(* IEC 61131-3 sources: volt/packages/volt-lsp-iec/test-corpus/awa-palletizer/Device/Plc Logic/Application/Library Manager/L_TS2P_TechModulesSynchronizingCamming, 208 files *)

(* ---- L_MB1P_CLUTCHDIRECTION.dut ---- *)
TYPE L_MB1P_CLUTCHDIRECTION :
(
	MCNEGATIVEDIRECTION := -1,
	MCCURRENTDIRECTION := 0,
	MCPOSITIVEDIRECTION := 1
);
END_TYPE

(* ---- L_MB1P_CLUTCHMODE.dut ---- *)
TYPE L_MB1P_CLUTCHMODE :
(
	ABSOLUTE := 0,
	RELATIVE := 1,
	RAMP_POS := 2,
	RAMP_TIME := 3,
	RAMP_SLAVE_DIST := 4,
	ABSOLUTE_IN_TARGET := 5,
	RAMP_VELACC := 6,
	DISTRELATIVE := 7
);
END_TYPE

(* ---- L_MB1P_STATES.dut ---- *)
TYPE L_MB1P_STATES :
(
	INIT := 1,
	READY := 2,
	HOMING := 3,
	JOGGING := 10,
	JOGPOS := 11,
	JOGNEG := 12,
	POSITION_TRIMMING := 20,
	TRIM_POS_PLUS := 21,
	TRIM_POS_MINUS := 22,
	SYNCPOS := 30,
	POS_IS_SYNCHRONISED := 31,
	POSITIONING_TO_START_POS := 32,
	SYNCSPEED := 40,
	SPEED_IS_SYNCHRONISED := 41,
	DECOUPLED_LOCAL_DRIVING := 50,
	CONTMOTION := 60,
	PREPARING_PATH := 61,
	CHECK_LIMITS := 62,
	SYNCLINEVEL := 70,
	CAMMING := 80,
	CAMMING_DONE := 81,
	CLUTCH_OPEN_INSTANT := 82,
	CLUTCH_CLOSE := 83,
	CLUTCH_OPEN := 84,
	CYCLICMOTION := 130,
	SETPARAMETERS := 140,
	CAMSEQUENCER_LOADCAMTABLE := 150,
	CAMSEQUENCER_CYCLICCAM1 := 151,
	CAMSEQUENCER_CYCLICCAM3 := 152,
	CAMSEQUENCER_CAM1CYCLICCAM3CAM1 := 153,
	CAMSEQUENCER_CAM1CAM2CYCLICCAM3CAM4CAM1 := 154,
	CALCULATION := 798,
	BUSY := 799,
	DONE := 800,
	EMERGENCYSTOP := 991,
	SLOWSTOP := 992,
	ABC := 993,
	STANDBY := 994,
	HALT := 995,
	STOP := 996,
	QUICKSTOP := 997,
	SERVICE := 998,
	ERROR := 999,
	SYSTEMFAULT := 1000
);
END_TYPE

(* ---- L_TF1P_STATES.dut ---- *)
TYPE L_TF1P_STATES :
(
	INIT := 1,
	READY := 2,
	HOMING := 3,
	JOGGING := 10,
	JOGPOS := 11,
	JOGNEG := 12,
	POSITION_TRIMMING := 20,
	TRIM_POS_PLUS := 21,
	TRIM_POS_MINUS := 22,
	SYNCPOS := 30,
	POS_IS_SYNCHRONISED := 31,
	POSITIONING_TO_START_POS := 32,
	SYNCSPEED := 40,
	SPEED_IS_SYNCHRONISED := 41,
	DECOUPLED_LOCAL_DRIVING := 50,
	CONTMOTION := 60,
	PREPARING_PATH := 61,
	CHECK_LIMITS := 62,
	SYNCLINEVEL := 70,
	CAMMING := 80,
	CAMMING_DONE := 81,
	CLUTCH_OPEN_INSTANT := 82,
	CLUTCH_CLOSE := 83,
	CLUTCH_OPEN := 84,
	CYCLICMOTION := 130,
	SETPARAMETERS := 140,
	CAMSEQUENCER_LOADCAMTABLE := 150,
	CAMSEQUENCER_CYCLICCAM1 := 151,
	CAMSEQUENCER_CYCLICCAM3 := 152,
	CAMSEQUENCER_CAM1CYCLICCAM3CAM1 := 153,
	CAMSEQUENCER_CAM1CAM2CYCLICCAM3CAM4CAM1 := 154,
	STANDBY := 994,
	HALT := 995,
	STOP := 996,
	QUICKSTOP := 997,
	SERVICE := 998,
	ERROR := 999
);
END_TYPE

(* ---- L_TF1P_SYNCMODE.dut ---- *)
TYPE L_TF1P_SYNCMODE :
(
	ABSOLUTE := 0,
	RELATIVE := 1,
	RAMP_TIME := 3,
	RAMP_VELACC := 4,
	RAMP_DIST := 5,
	DISTRELATIVE := 7
);
END_TYPE

(* ---- L_TS2M_SCDATA_FLYINGSAWSTATE.dut ---- *)
TYPE L_TS2M_SCDATA_FLYINGSAWSTATE :
STRUCT
	XEXECUTEMOVETOPARKPOS : BOOL;
	XMOVETOPARKPOSBUSY : BOOL;
	XMOVETOPARKPOSDONE : BOOL;
	XMOVETOPARKPOSABORTED : BOOL;
	EMOVETOPARKPOSDIRECTION : MC_DIRECTION := MC_DIRECTION.mcPositiveDirection;
	XPARKPOSREACHED : BOOL;
	XINPARKPOSITION : BOOL;
	XSTARTFLYINGSAW : BOOL;
	XFMFLYINGSAWPOSITIONING : BOOL;
	XFMFLYINGSAWINPOSITION : BOOL;
	XFMERROR : BOOL;
	EFMERRORID : L_IE1P_Error;
	EFM_STATE : L_TB2P_States;
	LRSETACCELERATION : LREAL;
	LRSETVELOCITY : LREAL;
	LRSETPOSITION : LREAL;
END_STRUCT
END_TYPE

(* ---- L_TS2M_SCDATA_FM_FLYINGSAW.dut ---- *)
TYPE L_TS2M_SCDATA_FM_FLYINGSAW :
STRUCT
	LRSTARTPOSOUT : LREAL;
	XGETNEXTMARK : BOOL;
	XRESETGETNEXTMARK : BOOL;
	XRESETMARKSTACK : BOOL;
	XNEWMARKRECEIVED : BOOL;
	XMARKSTACKEMPTY : BOOL;
	XMARKVALID : BOOL;
	LRMARKPOSOUT : LREAL;
	POSPROFILERCLUTCH_XENABLE : BOOL;
	POSPROFILERCLUTCH_XSYNCVEL : BOOL;
	POSPROFILERCLUTCH_XSYNCPOS : BOOL;
	POSPROFILERCLUTCH_XSYNCOUTINSTANT : BOOL;
	POSPROFILERCLUTCH_XMOVETOTARGETPOS : BOOL;
	POSPROFILERCLUTCH_LRTARGETPOS : LREAL;
	POSPROFILERCLUTCH_LRCORRECTTIMEBASE : LREAL;
	POSPROFILERCLUTCH_XEXECUTEGAP : BOOL;
	POSPROFILERCLUTCH_XAUXEXECUTEGAP : BOOL;
	POSPROFILERCLUTCH_LRCYCMASTERPOS : LREAL;
	POSPROFILERCLUTCH_LRCYCMASTERVEL : LREAL;
	POSPROFILERCLUTCH_LRCYCMASTERACC : LREAL;
	POSPROFILERCLUTCH_XERROR : BOOL;
	POSPROFILERCLUTCH_XBUSY : BOOL;
	POSPROFILERCLUTCH_XDONE : BOOL;
	POSPROFILERCLUTCH_XACCDECSYNC : BOOL;
	POSPROFILERCLUTCH_XVELSYNCHRONISED : BOOL;
	POSPROFILERCLUTCH_XPOSSYNCHRONISED : BOOL;
	POSPROFILERCLUTCH_XPOSITIONING : BOOL;
	POSPROFILERCLUTCH_XINPOSITION : BOOL;
	POSPROFILERCLUTCH_LRSETSLAVEPOSOUT : LREAL;
	POSPROFILERCLUTCH_LRSETSLAVEVELOUT : LREAL;
	POSPROFILERCLUTCH_LRSETSLAVEACCOUT : LREAL;
	POSPROFILERCLUTCH_XPROFILERESETTIMEVALID : BOOL;
	POSPROFILERCLUTCH_LRPROFILERESETTIME : LREAL;
	XMODECHANGE : BOOL;
	EFLYINGSAWMODE_OLD : L_TS2P_FlyingSawMode;
	LRACCDIST : LREAL;
	LRACCTIME : LREAL;
	XTPRECEIVED : BOOL;
	LRTPACTPOSITION : LREAL;
	XMASTERITFVALID : BOOL;
	BYMASTERID : POINTER TO BYTE;
	XMASTERITFVALID_LOCK : BOOL;
	BYMASTERID_LOCK : POINTER TO BYTE;
	XWARNING_TPRECPOSITIONNOTSUPPORTED : BOOL;
	LRSYNCOUTPOS : LREAL;
	XSTATESAWSYNCHRONIZED : BOOL;
	XSYNCOVERRIDEACTIVE : BOOL;
	XRAMPGENBUSY : BOOL;
	LRCUTLENGTHPROCESSED : LREAL;
	LRDISTTOCUTPOSITION : LREAL;
	LRMASTERPOS1 : LREAL;
	LRMASTERPOS2 : LREAL;
	LRSLAVEPOS1 : LREAL;
	LRSLAVEPOS2 : LREAL;
	LRCUTGAP_INT : LREAL;
	XHEADCUTDONE : BOOL;
	XMOVETOLOWERLIMITBUSY : BOOL;
	LRDIST_INT : LREAL;
	XTIMESYNCINVALID : BOOL;
	LRTIMESYNCIN_INT : LREAL;
	XWAITINGFORNEXTCUTBUSY : BOOL;
	XBALANCEDPROFILEACTIVE : BOOL;
	LRDISTTOTARGET : LREAL;
	LRFILTMATERIALVEL : LREAL;
	LRFILTMATERIALACC : LREAL;
	LRRESTTIMETARGETTOLOWERLIMIT : LREAL;
	FB_STACKCONTROLARRAYNOISE : L_MC1P_StackControlArray := STRUCT(iMaxLegth := 10);
	ALRDELTAVEL : ARRAY [0..10] OF LREAL;
	AXNOISE : ARRAY [0..5] OF BOOL;
	ALRVELTOLERANCE : ARRAY [0..5] OF LREAL;
	XNOISE : BOOL;
	XACCPOSITIV : BOOL;
	IACCCHANGEDIRECTIONCOUNTER : INT;
	LRVELTOLERANCE_INT : LREAL;
	LRMAXVELTOLERANCE : LREAL;
	LRMAXACCTOLERANCE : LREAL;
	LRCYCMASTERVEL : LREAL;
	LRCYCMASTERVEL_OLD : LREAL;
END_STRUCT
END_TYPE

(* ---- L_TS2P_CAMDATAXYVA.dut ---- *)
TYPE L_TS2P_CAMDATAXYVA :
STRUCT
	LRX : LREAL;
	LRY : LREAL;
	LRYS : LREAL;
	LRYSS : LREAL;
	LRYSSS : LREAL;
END_STRUCT
END_TYPE

(* ---- L_TS2P_CAMSEQUENCEMODE.dut ---- *)
TYPE L_TS2P_CAMSEQUENCEMODE :
(
	CYCLICCAM1 := 0,
	CYCLICCAM3 := 1,
	CAM1_CYCLICCAM3_CAM1 := 2,
	CAM1_CAM2_CYCLICCAM3_CAM4_CAM1 := 3
);
END_TYPE

(* ---- L_TS2P_CAMSTOPMODE.dut ---- *)
TYPE L_TS2P_CAMSTOPMODE :
(
	HALT := 0,
	MOVETOPARKPOS := 1
);
END_TYPE

(* ---- L_TS2P_CLUTCHINMODE.dut ---- *)
TYPE L_TS2P_CLUTCHINMODE :
(
	DISTABSOLUTE := 2,
	INSTANTABSOLUTE := 10
);
END_TYPE

(* ---- L_TS2P_CLUTCHOUTMODE.dut ---- *)
TYPE L_TS2P_CLUTCHOUTMODE :
(
	DISTABSOLUTE := 2,
	DISTRELATIVE := 3
);
END_TYPE

(* ---- L_TS2P_CORRECTIONMODE.dut ---- *)
TYPE L_TS2P_CORRECTIONMODE :
(
	POLYNOM5TH := 0,
	PROFILEGENERATOR := 1
);
END_TYPE

(* ---- L_TS2P_COUPLINGMODE.dut ---- *)
TYPE L_TS2P_COUPLINGMODE :
(
	UNITCOUPLING := 0,
	COUPLINGOVERCYCLELENGTH := 1
);
END_TYPE

(* ---- L_TS2P_CROSSCUTTERSTATEIN.dut ---- *)
TYPE L_TS2P_CROSSCUTTERSTATEIN :
STRUCT
	MASTERVALUES : L_MC1P_IAXIS_REF_MASTERVALUES;
	XEXECUTEMOVETOPARKPOS : BOOL;
	XSYNCIN : BOOL;
	XHOLDINPARKPOS : BOOL;
	LRPRODUCTLENGTH : LREAL;
	LROVERSPEED : LREAL;
	LRSETOFFSETPOSX : LREAL;
	XTRIMPOS : BOOL;
	XTRIMNEG : BOOL;
	XTRIMRESET : BOOL;
	SCTPRECDATA_MARKSENSOR : L_MC1P_TpReceiveData;
	SCTPRECDATA_TOOLSENSOR : L_MC1P_TpReceiveData;
	XTEACHMARKWINDOW : BOOL;
	XTEACHMARKWINDOWTOOL : BOOL;
	XGEARFACTORCORR : BOOL;
	XGEARFACTORCORRHOLD : BOOL;
END_STRUCT
END_TYPE

(* ---- L_TS2P_CROSSCUTTERSTATEOUT.dut ---- *)
TYPE L_TS2P_CROSSCUTTERSTATEOUT :
STRUCT
	XSYNCHRONISED : BOOL;
	XACCDECSYNC : BOOL;
	XOFFSETTRIMACTIVE : BOOL;
	XINPARKPOS : BOOL;
	XHOLDINPARKPOSACTIVE : BOOL;
	XCUTDONE : BOOL;
	XCUTTINGACTIVE : BOOL;
	LRACTCUTLENGTH : LREAL;
	LROFFSETTOTAL : LREAL;
	XTRQCTRLACTIVE : BOOL;
	LRSETMARKCORROUT : LREAL;
	XMARKWINDOWTEACHED : BOOL;
	LRGEARFACTORCORR : LREAL;
	LRSETTOOLCORROUT : LREAL;
	XMARKWINDOWTEACHEDTOOL : BOOL;
END_STRUCT
END_TYPE

(* ---- L_TS2P_CUTTINGMODEBASE.dut ---- *)
TYPE L_TS2P_CUTTINGMODEBASE :
(
	CUT_LENGTH := 0,
	FLOW_PACKER := 1
);
END_TYPE

(* ---- L_TS2P_CUTTINGMODESTATE.dut ---- *)
TYPE L_TS2P_CUTTINGMODESTATE :
(
	CUT_LENGTH := 0,
	FLOW_PACKER := 1,
	CUT_LENGTH_TP_CORRECTION := 2,
	CUT_ON_TP := 3
);
END_TYPE

(* ---- L_TS2P_ELECTRONICGEARBOXBASEIN.dut ---- *)
TYPE L_TS2P_ELECTRONICGEARBOXBASEIN :
STRUCT
	MASTERVALUES : L_MC1P_IAXIS_REF_MASTERVALUES;
	XSYNCIN : BOOL;
	LRSETBASEVEL : LREAL;
	LRSETOFFSETPOS : LREAL;
	LRSETOFFSETVEL : LREAL;
	XTRIMPOS : BOOL;
	XTRIMNEG : BOOL;
	XTRIMRESET : BOOL;
	XINVERTGEARFACTOR : BOOL;
END_STRUCT
END_TYPE

(* ---- L_TS2P_ELECTRONICGEARBOXBASEOUT.dut ---- *)
TYPE L_TS2P_ELECTRONICGEARBOXBASEOUT :
STRUCT
	XSYNCHRONISED : BOOL;
	XACCDECSYNC : BOOL;
	XOFFSETTRIMACTIVE : BOOL;
	XBASEVELOCITYACTIVE : BOOL;
	LROFFSETTOTALVEL : LREAL;
END_STRUCT
END_TYPE

(* ---- L_TS2P_FLEXCAMHIGHIN.dut ---- *)
TYPE L_TS2P_FLEXCAMHIGHIN :
STRUCT
	MASTERVALUES : L_MC1P_IAXIS_REF_MASTERVALUES;
	XCLUTCHCLOSE : BOOL;
	XLOADCLUTCHPOS : BOOL;
	LRLOADCLUTCHPOS : LREAL;
	XFINDCLUTCHXPOS : BOOL;
	XSYNCIN : BOOL;
	XSYNCPOSRESTORE : BOOL;
	XCAMCHANGEINSTANT : BOOL;
	LRSETOFFSETPOSX : LREAL;
	LRSETOFFSETPOSY : LREAL;
	LRSETSCALINGX : LREAL;
	LRSETSCALINGY : LREAL;
	CAMTABLE1 : MC_CAM_REF;
	CAMTABLE2 : MC_CAM_REF;
	CAMTABLE3 : MC_CAM_REF;
	CAMTABLE4 : MC_CAM_REF;
	WSETCAMTABLE : WORD := 1;
	XCAMSEQUENCER : BOOL;
END_STRUCT
END_TYPE

(* ---- L_TS2P_FLEXCAMHIGHOUT.dut ---- *)
TYPE L_TS2P_FLEXCAMHIGHOUT :
STRUCT
	XCLUTCHACTIVE : BOOL;
	XCLUTCHCLOSED : BOOL;
	XACCDECSYNC : BOOL;
	XSYNCHRONISED : BOOL;
	XMOVETOPARKPOSACTIVE : BOOL;
	XINPARKPOS : BOOL;
	XENDOFPROFILE : BOOL;
	LROFFSETPOSX : LREAL;
	LROFFSETPOSY : LREAL;
	LROFFSETSYNCPOS : LREAL;
	WACTIVECAMTABLE : WORD;
	XCAMSEQUENCERACTIVE : BOOL;
END_STRUCT
END_TYPE

(* ---- L_TS2P_FLEXCAMSTATEIN.dut ---- *)
TYPE L_TS2P_FLEXCAMSTATEIN :
STRUCT
	MASTERVALUES : L_MC1P_IAXIS_REF_MASTERVALUES;
	XSYNCIN : BOOL;
	XCAMCHANGEINSTANT : BOOL;
	LRSETOFFSETPOSX : LREAL;
	LRSETOFFSETPOSY : LREAL;
	LRSETSCALINGX : LREAL := 1;
	LRSETSCALINGY : LREAL := 1;
	CAMTABLE1 : MC_CAM_REF;
	CAMTABLE2 : MC_CAM_REF;
	CAMTABLE3 : MC_CAM_REF;
	CAMTABLE4 : MC_CAM_REF;
	WSETCAMTABLE : WORD := 1;
	XCAMSEQUENCER : BOOL;
END_STRUCT
END_TYPE

(* ---- L_TS2P_FLEXCAMSTATEOUT.dut ---- *)
TYPE L_TS2P_FLEXCAMSTATEOUT :
STRUCT
	XSYNCHRONISED : BOOL;
	XACCDECSYNC : BOOL;
	XCAMMINGBUSY : BOOL;
	XENDOFPROFILE : BOOL;
	LROFFSETPOSX : LREAL;
	LROFFSETPOSY : LREAL;
	WACTIVECAMTABLE : WORD;
	XCAMSEQUENCERACTIVE : BOOL;
END_STRUCT
END_TYPE

(* ---- L_TS2P_FLYINGSAWMODE.dut ---- *)
TYPE L_TS2P_FLYINGSAWMODE :
(
	MARKCONTROLLED := 0,
	LENGTHCONTROLLED := 1,
	LENGTHCONTROLLEDAUTOSYNC := 2
);
END_TYPE

(* ---- L_TS2P_FLYINGSAWPROFILEMODE.dut ---- *)
TYPE L_TS2P_FLYINGSAWPROFILEMODE :
(
	DEFAULT := 0,
	BALANCED := 1
);
END_TYPE

(* ---- L_TS2P_FLYINGSAWSTATEIN.dut ---- *)
TYPE L_TS2P_FLYINGSAWSTATEIN :
STRUCT
	MASTERVALUES : L_MC1P_IAXIS_REF_MASTERVALUES;
	XSTARTFLYINGSAW : BOOL;
	XSYNCININSTANT : BOOL;
	XEXECUTENEXTCUT : BOOL;
	XEXECUTEGAP : BOOL;
	XSETCUTTINGLENGTHINSTANT : BOOL;
	LRCUTTINGLENGTH : LREAL;
	LRSYNCOVERRIDE : LREAL := 1;
	XSETMATERIALCOUNTER : BOOL;
	XMOVETOPARKPOS : BOOL;
	XRESUMETARGETPOS : BOOL;
	XRESETMARKSTACK : BOOL;
	SCTPRECDATA_MARKSENSOR : L_MC1P.L_MC1P_TpReceiveData;
END_STRUCT
END_TYPE

(* ---- L_TS2P_FLYINGSAWSTATEOUT.dut ---- *)
TYPE L_TS2P_FLYINGSAWSTATEOUT :
STRUCT
	XSYNCHRONISED : BOOL;
	XACCDECSYNC : BOOL;
	XINPOSITION : BOOL;
	XPOSITIONING : BOOL;
	LRMATERIALCOUNTER : LREAL;
	LRTARGETPOS : LREAL;
	LRCUTGAP : LREAL;
	LRACTIVECUTTINGLENGTH : LREAL;
	WMARKSINSTACK : WORD;
END_STRUCT
END_TYPE

(* ---- L_TS2P_FLYINGSAWSTOPMODE.dut ---- *)
TYPE L_TS2P_FLYINGSAWSTOPMODE :
(
	HALT := 0,
	MOVETOPARKPOS := 1
);
END_TYPE

(* ---- L_TS2P_INTERFACEID.dut ---- *)
TYPE L_TS2P_INTERFACEID :
(
	L_TS2P_ISTRUCTPROVIDERFLYINGSAW := (L_TS2P_Internal.cdiEnumStartValue + 1),
	L_TS2P_ISTRUCTPROVIDERSYNCPOS := (L_TS2P_Internal.cdiEnumStartValue + 2),
	L_TS2P_ISTRUCTPROVIDERSYNCANDCORRECTION := (L_TS2P_Internal.cdiEnumStartValue + 3),
	L_TS2P_ISTRUCTPROVIDERFLEXCAMHIGH := (L_TS2P_Internal.cdiEnumStartValue + 4)
);
END_TYPE

(* ---- L_TS2P_OFFSETMODE.dut ---- *)
TYPE L_TS2P_OFFSETMODE :
(
	X_ZERO := 0,
	INSTANTABSOLUTE := 1,
	PROFGENABSOLUTE := 2
);
END_TYPE

(* ---- L_TS2P_SCALINGMODE.dut ---- *)
TYPE L_TS2P_SCALINGMODE :
(
	X_ZERO := 0,
	INSTANTABSOLUTE := 1,
	INSTANTRELATIVE := 2,
	PROFGENABSOLUTE := 3,
	PROFGENRELATIVE := 4
);
END_TYPE

(* ---- L_TS2P_SCAP_CROSSCUTTERBASE.dut ---- *)
TYPE L_TS2P_SCAP_CROSSCUTTERBASE :
STRUCT
END_STRUCT
END_TYPE

(* ---- L_TS2P_SCAP_CROSSCUTTERHIGH.dut ---- *)
TYPE L_TS2P_SCAP_CROSSCUTTERHIGH :
STRUCT
END_STRUCT
END_TYPE

(* ---- L_TS2P_SCAP_CROSSCUTTERSTATE.dut ---- *)
TYPE L_TS2P_SCAP_CROSSCUTTERSTATE :
STRUCT
END_STRUCT
END_TYPE

(* ---- L_TS2P_SCAP_ELECTRONICGEARBOXBASE.dut ---- *)
TYPE L_TS2P_SCAP_ELECTRONICGEARBOXBASE :
STRUCT
END_STRUCT
END_TYPE

(* ---- L_TS2P_SCAP_FLEXCAMHIGH.dut ---- *)
TYPE L_TS2P_SCAP_FLEXCAMHIGH :
STRUCT
END_STRUCT
END_TYPE

(* ---- L_TS2P_SCAP_FLEXCAMSTATE.dut ---- *)
TYPE L_TS2P_SCAP_FLEXCAMSTATE :
STRUCT
END_STRUCT
END_TYPE

(* ---- L_TS2P_SCAP_FLYINGSAWSTATE.dut ---- *)
TYPE L_TS2P_SCAP_FLYINGSAWSTATE :
STRUCT
END_STRUCT
END_TYPE

(* ---- L_TS2P_SCAP_SYNCANDCORRECTIONSTATE.dut ---- *)
TYPE L_TS2P_SCAP_SYNCANDCORRECTIONSTATE :
STRUCT
END_STRUCT
END_TYPE

(* ---- L_TS2P_SCAP_SYNCPOSBASE.dut ---- *)
TYPE L_TS2P_SCAP_SYNCPOSBASE :
STRUCT
END_STRUCT
END_TYPE

(* ---- L_TS2P_SCAP_TM_CROSSCUTTERBASE.dut ---- *)
TYPE L_TS2P_SCAP_TM_CROSSCUTTERBASE :
STRUCT
	AP_XENDOFPROFILEWINDOWSIZE : BOOL;
	AP_LRENDOFPROFILEWINDOWSIZE : LREAL := 0;
	AP_XOVERSPEEDUPPERLIMIT : BOOL;
	AP_LROVERSPEEDUPPERLIMIT : LREAL := 2;
	AP_XSETOFFSETSLAVE : BOOL;
	AP_LRSETOFFSETSLAVE : LREAL;
	AP_XOFFSETSLAVEPAR : BOOL;
	AP_LROFFSETSLAVEVEL : LREAL;
	AP_LROFFSETSLAVEACC : LREAL;
	AP_LROFFSETSLAVEDEC : LREAL;
	AP_LROFFSETSLAVEJERK : LREAL;
END_STRUCT
END_TYPE

(* ---- L_TS2P_SCAP_TM_CROSSCUTTERHIGH.dut ---- *)
TYPE L_TS2P_SCAP_TM_CROSSCUTTERHIGH :
STRUCT
END_STRUCT
END_TYPE

(* ---- L_TS2P_SCAP_TM_CROSSCUTTERSTATE.dut ---- *)
TYPE L_TS2P_SCAP_TM_CROSSCUTTERSTATE :
STRUCT
	AP_XTPAXISDELAYCYCLE : BOOL;
	AP_LRTPAXISDELAYCYCLE : LREAL;
	AP_XTPAXISCOMPFACTOR : BOOL;
	AP_LRTPAXISCOMPFACTOR : LREAL;
	AP_XUPPERCORRPOS : BOOL;
	AP_LRUPPERCORRPOS : LREAL;
	AP_XLOWERCORRPOS : BOOL;
	AP_LRLOWERCORRPOS : LREAL;
	AP_XCUTTINGANGLESTOPCAM : BOOL;
	AP_LRCUTTINGANGLESTOPCAM : LREAL := 10;
	AP_XSETCUTLENGTHINPRODUCT : BOOL;
END_STRUCT
END_TYPE

(* ---- L_TS2P_SCAP_TM_ELECTRONICGEARBOXBASE.dut ---- *)
TYPE L_TS2P_SCAP_TM_ELECTRONICGEARBOXBASE :
STRUCT
	AP_XGEARINGNUMERATOR : BOOL;
	AP_DWGEARINGNUMERATOR : DWORD := 1;
	AP_XGEARINGDENOMINATOR : BOOL;
	AP_DWGEARINGDENOMINATOR : DWORD := 1;
	AP_XLIMITALLOWEDDIRECTION : BOOL;
	AP_LREXTTHRESHOLDDIRECTION : LREAL;
END_STRUCT
END_TYPE

(* ---- L_TS2P_SCAP_TM_FLEXCAM.dut ---- *)
TYPE L_TS2P_SCAP_TM_FLEXCAM :
STRUCT
	AP_LREXTTHRESHOLDDIRECTION : LREAL;
	AP_LRMASTERVELSTANDSTILLDEADBAND : LREAL;
	AP_XENDOFPROFILEWINDOWSIZE : BOOL;
	AP_LRENDOFPROFILEWINDOWSIZE : LREAL;
	AP_XSETVALUEMODE : BOOL;
	AP_ESETVALUEMODE : L_MC1P_SetValueMode := L_MC1P_SetValueMode.PosVelAcc;
END_STRUCT
END_TYPE

(* ---- L_TS2P_SCAP_TM_FLEXCAMBASE.dut ---- *)
TYPE L_TS2P_SCAP_TM_FLEXCAMBASE :
STRUCT
	AP_XENDOFPROFILEWINDOWSIZE : BOOL;
	AP_LRENDOFPROFILEWINDOWSIZE : LREAL := 0;
	AP_XCALCAMPROFILER : BOOL := TRUE;
	AP_XSETVALUEMODE : BOOL;
	AP_ESETVALUEMODE : L_MC1P_SetValueMode := L_MC1P_SetValueMode.PosVelAcc;
END_STRUCT
END_TYPE

(* ---- L_TS2P_SCAP_TM_FLEXCAMSTATE.dut ---- *)
TYPE L_TS2P_SCAP_TM_FLEXCAMSTATE :
STRUCT
END_STRUCT
END_TYPE

(* ---- L_TS2P_SCAP_TM_FLYINGSAWSTATE.dut ---- *)
TYPE L_TS2P_SCAP_TM_FLYINGSAWSTATE :
STRUCT
	AP_XLOADTOTALCUTTINGLENGTH : BOOL;
	AP_LRLOADTOTALCUTTINGLENGTH : LREAL;
	AP_XLOADTARGETPOS : BOOL;
	AP_LRLOADTARGETPOS : LREAL;
	AP_XRANGEOFTOLERANCE : BOOL;
	AP_LRRANGEOFTOLERANCE : LREAL;
	AP_XMARKDETECTERRCOMP : BOOL;
	AP_LRMARKDETECTERRCOMP : LREAL;
	AP_XTASKCYCLEDELAY : BOOL;
	AP_BYTASKCYCLEDELAY : BYTE;
END_STRUCT
END_TYPE

(* ---- L_TS2P_SCAP_TM_SYNCANDCORRECTIONSTATE.dut ---- *)
TYPE L_TS2P_SCAP_TM_SYNCANDCORRECTIONSTATE :
STRUCT
	AP_DIDEADTIMECOMP : DINT;
END_STRUCT
END_TYPE

(* ---- L_TS2P_SCAP_TM_SYNCPOSBASE.dut ---- *)
TYPE L_TS2P_SCAP_TM_SYNCPOSBASE :
STRUCT
	AP_XLOADGEARBOXPOSOUT : BOOL;
	AP_LRLOADGEARBOXPOSOUT : LREAL;
	AP_XLOADTRIMOFFSET : BOOL;
	AP_LRLOADTRIMOFFSET : LREAL;
	AP_XLOADOFFSETSYNC : BOOL;
	AP_LRLOADOFFSETSYNC : LREAL;
	AP_XLIMITALLOWEDDIRECTION : BOOL;
	AP_LREXTTHRESHOLDDIRECTION : LREAL;
	AP_LRMASTERVELSTANDSTILLDEADBAND : LREAL;
END_STRUCT
END_TYPE

(* ---- L_TS2P_SCDATA_TM_FLEXCAM.dut ---- *)
TYPE L_TS2P_SCDATA_TM_FLEXCAM :
STRUCT
	XEXECUTEMOVETOPARKPOS : BOOL;
	XHALTFLEXCAM : BOOL;
	XMOVETOPARKPOSBUSY : BOOL;
	XMOVETOPARKPOSABORTED : BOOL;
	MASTERVALUES_ITFVALID : L_MC1P_IAXIS_REF_MASTERVALUES;
	LRMASTERPOS_OLD : LREAL;
	LRMASTERVEL_OLD : LREAL;
	LRSETPOSITIONFORSYNCMASTER : LREAL;
	LRSETVELOCITYFORSYNCMASTER : LREAL;
	LRSETACCELERATIONFORSYNCMASTER : LREAL;
	LRCYCLELENGTHMASTER : LREAL;
	ETRAVERSINGRANGEMASTER : L_MC1P_TraversingRange;
	LRSETPOSITIONAXIS : LREAL;
	LRSETVELOCITYAXIS : LREAL;
	LRSETACCELERATIONAXIS : LREAL;
	WACTDIRECTIONMASTER : WORD;
	XCAMSEQUENCERERROR : BOOL;
	ECAMSEQUENCERERROR : L_IE1P_Error;
	XCAMERROR : BOOL;
	ECAMERROR : L_IE1P_Error;
	XCAMBUSY : BOOL;
	XCAMDONE : BOOL;
	XLOCKTOCAMRESTORE : BOOL;
	ESYNCINMODE : L_TS2P_SyncInMode := L_TS2P_SyncInMode.ProfGenAbsolute;
	XCLUTCHBUSY : BOOL;
	XCLUTCHDONE : BOOL;
	XCLUTCHACCDECSYNCLED : BOOL;
	LRSETCLUTCHPOSOUT : LREAL;
	LRSETCLUTCHVELOUT : LREAL;
	LRSETCLUTCHACCOUT : LREAL;
	LRSETCLUTCHPOSOUTOLD : LREAL;
	LRSETCLUTCHVELOUTOLD : LREAL;
	XCLUTCHERROR : BOOL;
	ECLUTCHERROR : L_IE1P_Error;
	XENABLEALLOWEDDIRECTION : BOOL;
	LRALLOWEDDIRECTIONSETPOSOUT : LREAL;
	LRALLOWEDDIRECTIONSETVELOUT : LREAL;
	LRALLOWEDDIRECTIONSETACCOUT : LREAL;
	XALLOWEDDIRECTIONERROR : BOOL;
	XALLOWEDDIRECTIONWARNING : BOOL;
	EALLOWEDDIRECTIONERROR : L_IE1P_Error;
	XPOSFOLLOWERENABLE : BOOL;
	XPOSFOLLOWERBUSY : BOOL;
	XENABLETRANSSYNCHRONISED : BOOL;
	LRTASKCYCLE : LREAL;
	XLOCKTOCAM : BOOL;
	XCAMCHANGEINSTANT_INT : BOOL;
	LRSETOFFSETMASTER_INT : LREAL;
	LRSETOFFSETSLAVE_INT : LREAL;
	LRSETSCALINGMASTER_INT : LREAL := 1;
	LRSETSCALINGSLAVE_INT : LREAL := 1;
	SCPAR_INT : L_TS2P_scPar_TM_FlexCam;
	XLOCKTOCAMERROR : BOOL;
	ELOCKTOCAMERROR : L_IE1P_Error;
	XCAMTABLEVALID : BOOL;
	XCAMMINGBUSY : BOOL;
	XLOCKTOCAMDONE : BOOL;
	XLOCKTOCAMBUSY : BOOL;
	XLOCKTOCAMBUSYLED : BOOL;
	XLOCKTOCAMBUSYGENERAL : BOOL;
	EPOSFOLLOWERMODE : L_MC1P_SetValueMode;
	XLOADCAMXVALUEBUSY : BOOL;
	XDIRECTIONLIMITED : BOOL;
	XFINDCLUTCHXPOS : BOOL;
	XVISULAMPFALSE : BOOL;
	LRSETVELOLD : LREAL;
END_STRUCT
END_TYPE

(* ---- L_TS2P_SCDATA_TM_SYNCANDCORRECTIONSTATE.dut ---- *)
TYPE L_TS2P_SCDATA_TM_SYNCANDCORRECTIONSTATE :
STRUCT
	MASTERVALUES_ITFVALID : L_MC1P_IAXIS_REF_MASTERVALUES;
	XMASTERITFVALID : BOOL;
	XMASTERVALUECORRENABLED : BOOL;
	LRSETPOSOLD : LREAL;
	LRMASTERSETPOSOLD : LREAL;
	LRMASTERACTPOSITIONOLD : LREAL;
	LRSETVELOCITYGEARING : LREAL;
	LRSENSORSETPOS : LREAL;
	XMARKDISTCHANGED : BOOL;
	LRACTOFFSETMASTER : LREAL;
	LRACTOFFSETSLAVE : LREAL;
	LRLOWERCORRPOS : LREAL;
	LRUPPERCORRPOS : LREAL;
	LRMARKDIST : LREAL;
	LRACTOFFSETX : LREAL;
	XVALUESTORED : BOOL;
	XFIRSTVALUESTORED : BOOL;
	XTEACHTPSENSOROLD : BOOL;
	XTPSENSORTEACHEDOLD : BOOL;
	LRMARKSTACKLENGTH : LREAL;
	DWACTTIMESTAMPMARKWINDOW : DWORD;
	DWRECTIMESTAMPMARKWINDOW : DWORD;
	XVALUESTOREDMARKWINDOW : BOOL;
	XSUPPORTTIMESTAMPMARKWINDOW : BOOL;
	XVALUESTOREDMARKSTACK : BOOL;
	DWACTTIMESTAMPMARKSTACK : DWORD;
	DWRECTIMESTAMPMARKSTACK : DWORD;
	XVALUESTOREDTPCONVERTER : BOOL;
	LRTPACTPOSITIONTPCONVERTER : LREAL;
	LRACTMARKDIST : LREAL;
	LRMARKDISTINTEGRATOR : LREAL;
	LRTPDEADTIMEDIFF : LREAL;
	LRMARKERROR : LREAL;
	LRMARKERRORLIMITED : LREAL;
	LRMARKERRORGEARFACTOR : LREAL;
	LRCORRRESIDUAL : LREAL;
	LRDELTAGEARFACTORCORR : LREAL;
	LRGEARFACTORINTEGRATOR : LREAL;
	LRGEARFACTORNUMERATOR : LREAL;
	LRGEARFACTORNUMERATORCORR : LREAL;
	LRGEARFACTORDENOMINATOR : LREAL;
	LRGEARFACTORNUMERATORCORRLIMITED : LREAL;
	LRSTARTPOS : LREAL;
	ECORRMODEMASTEROLD : L_TS2P_CorrectionMode;
	LRSETVELOUTCORRECTION : LREAL;
	LRSETPOSOUTCORRECTION : LREAL;
	XVALUESTOREDCORRMARKERROR : BOOL;
END_STRUCT
END_TYPE

(* ---- L_TS2P_SCDATA_TM_SYNCPOSBASE.dut ---- *)
TYPE L_TS2P_SCDATA_TM_SYNCPOSBASE :
STRUCT
	MASTERVALUES_ITFVALID : L_MC1P_IAXIS_REF_MASTERVALUES;
	XHOMINGNOTNEEDED : BOOL;
	LRSETPOSITIONFORSYNCMASTER : LREAL;
	LRSETVELOCITYFORSYNCMASTER : LREAL;
	LRSETACCELERATIONFORSYNCMASTER : LREAL;
	LRCYCLELENGTHMASTER : LREAL;
	ETRAVERSINGRANGEMASTER : L_MC1P_TraversingRange;
	WACTDIRECTIONMASTER : WORD;
	XOFFSETTRIMERROR : BOOL;
	EOFFSETTRIMERROR : L_IE1P_Error;
	XADDOFFSETERROR : BOOL;
	EADDOFFSETERROR : L_IE1P_Error;
	LROFFSETAXISCONVERTER : LREAL;
	WTRAVERSINGRANGECOMBINATION : WORD;
	WTRAVERSINGRANGECOMBINATIONOLD : WORD;
	XGEARBOXERROR : BOOL;
	EGEARBOXERROR : L_IE1P_Error;
	LRBASEVELLIMITED : LREAL;
	XCLUTCHENABLE : BOOL;
	XCLUTCHSYNCIN : BOOL;
	XCLUTCHSYNCPOSRESTORE : BOOL;
	LRSETVELCLUTCHOFFSET : LREAL;
	LRSETACCCLUTCHOFFSET : LREAL;
	LRSETDECCLUTCHOFFSET : LREAL;
	LRSETJERKCLUTCHOFFSET : LREAL;
	ESYNCMODE : L_TB2P_SyncMode := L_TB2P_SyncMode.ProfGenAbsolute;
	XCLUTCHBUSY : BOOL;
	XCLUTCHDONE : BOOL;
	XCLUTCHSYNCHRONISED : BOOL;
	XCLUTCHACCDECSYNC : BOOL;
	LRCLUTCHSETPOSOUT : LREAL;
	LRCLUTCHSETVELOUT : LREAL;
	LRCLUTCHSETACCOUT : LREAL;
	LRSYNCOFFSET : LREAL;
	XCLUTCHERROR : BOOL;
	ECLUTCHERROR : L_IE1P_Error;
	LRALLOWEDDIRECTIONSETPOSOUT : LREAL;
	LRALLOWEDDIRECTIONSETVELOUT : LREAL;
	LRALLOWEDDIRECTIONSETACCOUT : LREAL;
	XALLOWEDDIRECTIONERROR : BOOL;
	XALLOWEDDIRECTIONWARNING : BOOL;
	EALLOWEDDIRECTIONERROR : L_IE1P_Error;
	XPOSFOLLOWERENABLE : BOOL;
	LRPOSFOLLOWERSETPOSIN : LREAL;
	LRPOSFOLLOWERSETVELIN : LREAL;
	XENABLETRANSBASEVEL : BOOL;
	XENABLETRANSSYNCHRONISED : BOOL;
	XENABLEOLD : BOOL;
	LRTASKCYCLE : LREAL;
	LRCYCLELENGTH : LREAL;
	ETRAVERSINGRANGE : L_MC1P_TraversingRange;
	LRSETPOSITION : LREAL;
	LRSETVELOCITY : LREAL;
	LRSETACCELERATION : LREAL;
	XREQUESTTOSTANDBY : BOOL;
END_STRUCT
END_TYPE

(* ---- L_TS2P_SCERRORINFO.dut ---- *)
TYPE L_TS2P_SCERRORINFO :
STRUCT
	XERROR : BOOL;
	XWARNING : BOOL;
	EERRORID : L_IE1P_Error;
	XAXISERROR : BOOL;
	XAXISWARNING : BOOL;
	EAXISERRORID : L_IE1P_Error;
	XDRIVEERROR : BOOL;
	XDRIVEWARNING : BOOL;
	DWDRIVEERRORID : DWORD;
END_STRUCT
END_TYPE

(* ---- L_TS2P_SCPAR_CROSSCUTTERBASE.dut ---- *)
TYPE L_TS2P_SCPAR_CROSSCUTTERBASE :
STRUCT
END_STRUCT
END_TYPE

(* ---- L_TS2P_SCPAR_CROSSCUTTERSTATE.dut ---- *)
TYPE L_TS2P_SCPAR_CROSSCUTTERSTATE :
STRUCT
END_STRUCT
END_TYPE

(* ---- L_TS2P_SCPAR_ELECTRONICGEARBOXBASE.dut ---- *)
TYPE L_TS2P_SCPAR_ELECTRONICGEARBOXBASE :
STRUCT
END_STRUCT
END_TYPE

(* ---- L_TS2P_SCPAR_FLEXCAMHIGH.dut ---- *)
TYPE L_TS2P_SCPAR_FLEXCAMHIGH :
STRUCT
END_STRUCT
END_TYPE

(* ---- L_TS2P_SCPAR_FLEXCAMSTATE.dut ---- *)
TYPE L_TS2P_SCPAR_FLEXCAMSTATE :
STRUCT
END_STRUCT
END_TYPE

(* ---- L_TS2P_SCPAR_FLYINGSAWSTATE.dut ---- *)
TYPE L_TS2P_SCPAR_FLYINGSAWSTATE :
STRUCT
END_STRUCT
END_TYPE

(* ---- L_TS2P_SCPAR_SYNCANDCORRECTIONSTATE.dut ---- *)
TYPE L_TS2P_SCPAR_SYNCANDCORRECTIONSTATE :
STRUCT
END_STRUCT
END_TYPE

(* ---- L_TS2P_SCPAR_SYNCPOSBASE.dut ---- *)
TYPE L_TS2P_SCPAR_SYNCPOSBASE :
STRUCT
END_STRUCT
END_TYPE

(* ---- L_TS2P_SCPAR_TM_CROSSCUTTERBASE.dut ---- *)
TYPE L_TS2P_SCPAR_TM_CROSSCUTTERBASE :
STRUCT
	LRSETOFFSETTRIMVEL : LREAL := 10.0;
	LRSETOFFSETTRIMACC : LREAL := 100.0;
	LRSETOFFSETTRIMDEC : LREAL := 100.0;
	LRSETOFFSETTRIMJERK : LREAL := 10000.0;
	ETRIMMODE : L_TS2P_TrimMode := L_TS2P_TrimMode.position;
	LRTRIMDIST : LREAL := 1;
	ESYNCMODE : L_TS2P_SyncModeCrossCutter;
	LRMASTERSYNCINDIST : LREAL := 0;
	LRMASTERSYNCOUTDIST : LREAL := 0;
	XMASTERABSOLUTE : BOOL := TRUE;
	LRSTARTXPOSRELATIVE : LREAL := 0;
	BYSTARTTOOLNO : BYTE := 0;
	BYNUMOFTOOLS : BYTE := 1;
	LRCUTTINGANGLE : LREAL := 10;
	LRTOOLCIRCUMFERENCE : LREAL := 75.55555;
	XCALCCAMBOUNDS : BOOL := FALSE;
	LRMASTERMAXVEL : LREAL := 100;
	LRMASTERMAXACC : LREAL := 1000;
	LRSCALINGMASTER : LREAL := 1;
	EPROFILETYPE : L_MC2P_LawOfMotion := L_MC2P_LawOfMotion.Poly5;
END_STRUCT
END_TYPE

(* ---- L_TS2P_SCPAR_TM_CROSSCUTTERBASEEXTENSION.dut ---- *)
TYPE L_TS2P_SCPAR_TM_CROSSCUTTERBASEEXTENSION :
STRUCT
	ECUTTINGMODE : L_TS2P_CuttingModeBase := L_TS2P_CuttingModeBase.cut_length;
END_STRUCT
END_TYPE

(* ---- L_TS2P_SCPAR_TM_CROSSCUTTERHIGH.dut ---- *)
TYPE L_TS2P_SCPAR_TM_CROSSCUTTERHIGH :
STRUCT
END_STRUCT
END_TYPE

(* ---- L_TS2P_SCPAR_TM_CROSSCUTTERSTATE.dut ---- *)
TYPE L_TS2P_SCPAR_TM_CROSSCUTTERSTATE :
STRUCT
	ECUTTINGMODE : L_TS2P_CuttingModeState;
	ALRCUTLENGTHINPRODUCT : ARRAY [1..10] OF LREAL;
	LRMINPRODUCTLENGTH : LREAL := 50;
	LRTRQCTRLGAIN : LREAL := 0;
	LRTRQCTRLRATETIME : LREAL := 0;
	LRMINERTIA : LREAL := 0;
	XCORRMARKERRORMASTER : BOOL := TRUE;
	LRSENSORTOOLDISTMASTER : LREAL := 0.0;
	LRMAXCORRPOSMASTER : LREAL := 30.0;
	LRMAXCORRNEGMASTER : LREAL := -30.0;
	XENABLEMARKWINDOWMASTER : BOOL;
	LRMARKWINDOWSIZEMASTER : LREAL := 90.0;
	LRSETOFFSETMARKWINDOWMASTER : LREAL := 0.0;
	LRGEARFACTORCORRGAINMASTER : LREAL := 0.1;
	LRMAXGEARFACTORCORRMASTER : LREAL := 10;
	DWMAXNUMBERVIRTUALMARKSMASTER : DWORD := 5;
	XLOADREGPOS : BOOL;
	LRLOADREGPOS : LREAL;
	XCALCTOOLERROR : BOOL := FALSE;
	XCORRTOOLERROR : BOOL := TRUE;
	LRSENSORTOOLDISTTOOL : LREAL := 0.0;
	XENABLEMARKWINDOWTOOL : BOOL := FALSE;
	LRMAXCORRPOSTOOL : LREAL := 30.0;
	LRMAXCORRNEGTOOL : LREAL := -30.0;
	LRUPPERCORRPOSTOOL : LREAL := 180.0;
	LRLOWERCORRPOSTOOL : LREAL := 90.0;
	LRMARKWINDOWSIZETOOL : LREAL := 90.0;
	LRSETOFFSETMARKWINDOWTOOL : LREAL := 0.0;
	DWMAXNUMBERVIRTUALMARKSTOOL : DWORD := 5;
END_STRUCT
END_TYPE

(* ---- L_TS2P_SCPAR_TM_ELECTRONICGEARBOXBASE.dut ---- *)
TYPE L_TS2P_SCPAR_TM_ELECTRONICGEARBOXBASE :
STRUCT
	ECOUPLINGMODE : L_TS2P_CouplingMode := 1;
	LRTOLERANCEINVERTGEARFACTOR : LREAL := 0;
END_STRUCT
END_TYPE

(* ---- L_TS2P_SCPAR_TM_FLEXCAM.dut ---- *)
TYPE L_TS2P_SCPAR_TM_FLEXCAM :
STRUCT
	ECLUTCHINMODE : L_TS2P_ClutchInMode := L_TS2P_ClutchInMode.DistAbsolute;
	ECLUTCHOUTMODE : L_TS2P_ClutchOutMode := L_TS2P_ClutchOutMode.DistAbsolute;
	LRCLUTCHINDISTX : LREAL := 90.0;
	LRCLUTCHOUTDISTX : LREAL := 90.0;
	LRCLUTCHOUTPOSX : LREAL := 0;
	XCAMCYCLIC : BOOL := TRUE;
	XMASTERABSOLUTE : BOOL := TRUE;
	XSLAVEABSOLUTE : BOOL := TRUE;
	EOFFSETMODEX : L_TS2P_OffsetMode := L_TS2P_OffsetMode.x_zero;
	EOFFSETMODEY : L_TS2P_OffsetMode := L_TS2P_OffsetMode.x_zero;
	LRSETOFFSETSCALINGXVEL : LREAL := 100.0;
	LRSETOFFSETSCALINGXACC : LREAL := 1000.0;
	LRSETOFFSETSCALINGXDEC : LREAL := 1000.0;
	LRSETOFFSETSCALINGXJERK : LREAL := 1000000.0;
	ESCALINGMODEX : L_TS2P_ScalingMode := L_TS2P_ScalingMode.x_zero;
	ESCALINGMODEY : L_TS2P_ScalingMode := L_TS2P_ScalingMode.x_zero;
	LRSETOFFSETSCALINGYVEL : LREAL := 100.0;
	LRSETOFFSETSCALINGYACC : LREAL := 1000.0;
	LRSETOFFSETSCALINGYDEC : LREAL := 1000.0;
	LRSETOFFSETSCALINGYJERK : LREAL := 1000000.0;
	XCALCCAMBOUNDS : BOOL;
	LRMASTERMAXVEL : LREAL := 100;
	LRMASTERMAXACC : LREAL := 1000;
	ECAMSEQUENCEMODE : L_TS2P_CamSequenceMode := L_TS2P_CamSequenceMode.CyclicCam1;
	ESYNCINMODE : L_TS2P_SyncInMode := L_TS2P_SyncInMode.ProfGenAbsolute;
	ESYNCOUTMODE : L_TS2P_CamStopMode := L_TS2P_CamStopMode.Halt;
	ESYNCDIRECTION : L_TS2P_SyncDirection := L_TS2P_SyncDirection.PositiveDirection;
	LRSYNCVEL : LREAL := 100;
	LRSYNCACC : LREAL := 1000.0;
	LRSYNCDEC : LREAL := 1000.0;
	LRSYNCJERK : LREAL := 1000000.0;
	LRPARKPOSITION : LREAL := 0.0;
	EALLOWEDDIRECTION : L_TB2P_AllowedDirection := L_TB2P_AllowedDirection.both;
	XLIMITALLOWEDDIRECTION : BOOL := FALSE;
	LRTOLERANCEALLOWEDDIRECTION : LREAL := 5;
END_STRUCT
END_TYPE

(* ---- L_TS2P_SCPAR_TM_FLEXCAMBASE.dut ---- *)
TYPE L_TS2P_SCPAR_TM_FLEXCAMBASE :
STRUCT
	ESYNCMODE : L_TS2P_SyncModeFlexCam := L_TS2P_SyncModeFlexCam.ProfGenAbsolute;
	EALLOWEDDIRECTION : L_TB2P_AllowedDirection := L_TB2P_AllowedDirection.both;
	LRMASTERSYNCINDIST : LREAL := 100;
	LRMASTERSYNCINPOS : LREAL := 0;
	LRMASTERSYNCOUTDIST : LREAL := 100;
	LRSLAVESYNCOUTPOS : LREAL := 0;
	LRSYNCVEL : LREAL := 100;
	LRSYNCACC : LREAL := 1000.0;
	LRSYNCDEC : LREAL := 1000.0;
	LRSYNCJERK : LREAL := 1000000.0;
	XCAMCYCLIC : BOOL := TRUE;
	XMASTERABSOLUTE : BOOL := TRUE;
	XSLAVEABSOLUTE : BOOL := TRUE;
	EOFFSETMODEX : L_TS2P_OffsetMode := L_TS2P_OffsetMode.x_zero;
	EOFFSETMODEY : L_TS2P_OffsetMode := L_TS2P_OffsetMode.x_zero;
	LRSETOFFSETSCALINGXVEL : LREAL := 100.0;
	LRSETOFFSETSCALINGXACC : LREAL := 1000.0;
	LRSETOFFSETSCALINGXDEC : LREAL := 1000.0;
	LRSETOFFSETSCALINGXJERK : LREAL := 1000000.0;
	ESCALINGMODEX : L_TS2P_ScalingMode := L_TS2P_ScalingMode.x_zero;
	ESCALINGMODEY : L_TS2P_ScalingMode := L_TS2P_ScalingMode.x_zero;
	LRSETOFFSETSCALINGYVEL : LREAL := 100.0;
	LRSETOFFSETSCALINGYACC : LREAL := 1000.0;
	LRSETOFFSETSCALINGYDEC : LREAL := 1000.0;
	LRSETOFFSETSCALINGYJERK : LREAL := 1000000.0;
	XCALCCAMBOUNDS : BOOL;
	LRMASTERMAXVEL : LREAL := 100;
	LRMASTERMAXACC : LREAL := 1000;
END_STRUCT
END_TYPE

(* ---- L_TS2P_SCPAR_TM_FLEXCAMSTATE.dut ---- *)
TYPE L_TS2P_SCPAR_TM_FLEXCAMSTATE :
STRUCT
	ECAMSEQUENCEMODE : L_TS2P_CamSequenceMode := L_TS2P_CamSequenceMode.CyclicCam1;
END_STRUCT
END_TYPE

(* ---- L_TS2P_SCPAR_TM_FLYINGSAWSTATE.dut ---- *)
TYPE L_TS2P_SCPAR_TM_FLYINGSAWSTATE :
STRUCT
	LRSYNCVEL : LREAL := 100;
	LRSYNCACC : LREAL := 1000.0;
	LRSYNCDEC : LREAL := 1000.0;
	LRSYNCJERK : LREAL := 1000000.0;
	LRSETMATERIALPOS : LREAL := 0;
	LRUPPERLIMIT : LREAL := 1000;
	LRLOWERLIMIT : LREAL := 0;
	LRGAP : LREAL;
	LRBLADEWIDTH : LREAL := 0;
	EPROFILEMODE : L_TS2P_FlyingSawProfileMode := L_TS2P_FlyingSawProfileMode.Default;
	EFLYINGSAWMODE : L_TS2P_FlyingSawMode := L_TS2P_FlyingSawMode.MarkControlled;
	EFLYINGSAWSTOPMODE : L_TS2P_FlyingSawStopMode := L_TS2P_FlyingSawStopMode.Halt;
	LRPARKPOSITION : LREAL := 0;
	LRMARKSENSORPOS : LREAL;
	XPOSINWINDOW : BOOL;
	LRTOLERANCEPOSINWINDOW : LREAL;
	LRDWELLTIMEPOSINWINDOW : LREAL := 0.05;
	LRTOLERANCEMASTERVELINWINDOW : LREAL;
END_STRUCT
END_TYPE

(* ---- L_TS2P_SCPAR_TM_SYNCANDCORRECTIONSTATE.dut ---- *)
TYPE L_TS2P_SCPAR_TM_SYNCANDCORRECTIONSTATE :
STRUCT
	ESOURCEFORCORRWINDOW : L_TS2P_SourceForCorrWindow := L_TS2P_SourceForCorrWindow.Slave;
	XCALCMARKERRORMASTER : BOOL := FALSE;
	XCORRMARKERRORMASTER : BOOL := TRUE;
	LRSENSORTOOLDISTMASTER : LREAL := 0.0;
	LRMARKDISTMASTER : LREAL := 360.0;
	ECORRMODEMASTER : L_TS2P_CorrectionMode := L_TS2P_CorrectionMode.Polynom5th;
	LRCORRVELMASTER : LREAL := 100;
	LRCORRACCMASTER : LREAL := 100;
	LRCORRDECMASTER : LREAL := 100;
	LRCORRJERKMASTER : LREAL := 10000;
	LRMAXCORRPOSMASTER : LREAL := 30.0;
	LRMAXCORRNEGMASTER : LREAL := -30.0;
	LRUPPERCORRPOSMASTER : LREAL := 180.0;
	LRLOWERCORRPOSMASTER : LREAL := 90.0;
	XENABLEMARKWINDOWMASTER : BOOL;
	LRMARKWINDOWSIZEMASTER : LREAL := 90.0;
	LRSETOFFSETMARKWINDOWMASTER : LREAL := 0.0;
	LRGEARFACTORCORRGAINMASTER : LREAL := 0.1;
	LRMAXGEARFACTORCORRMASTER : LREAL := 10;
	DWMAXNUMBERVIRTUALMARKSMASTER : DWORD := 5;
	XCALCTOOLERROR : BOOL := FALSE;
	XCORRTOOLERROR : BOOL := TRUE;
	LRSENSORTOOLDISTTOOL : LREAL := 0.0;
	LRMAXCORRPOSTOOL : LREAL := 30.0;
	LRMAXCORRNEGTOOL : LREAL := -30.0;
	ECORRMODETOOL : L_TS2P_CorrectionMode := L_TS2P_CorrectionMode.Polynom5th;
	LRCORRVELTOOL : LREAL := 100;
	LRCORRACCTOOL : LREAL := 100;
	LRCORRDECTOOL : LREAL := 100;
	LRCORRJERKTOOL : LREAL := 10000;
	LRUPPERCORRPOSTOOL : LREAL := 180.0;
	LRLOWERCORRPOSTOOL : LREAL := 90.0;
	XENABLEMARKWINDOWTOOL : BOOL := FALSE;
	LRMARKWINDOWSIZETOOL : LREAL := 90.0;
	LRSETOFFSETMARKWINDOWTOOL : LREAL := 0.0;
	DWMAXNUMBERVIRTUALMARKSTOOL : DWORD := 5;
	XLOADREGPOS : BOOL;
	LRLOADREGPOS : LREAL;
END_STRUCT
END_TYPE

(* ---- L_TS2P_SCPAR_TM_SYNCPOSBASE.dut ---- *)
TYPE L_TS2P_SCPAR_TM_SYNCPOSBASE :
STRUCT
	ESYNCMODE : L_TB2P_SyncMode := L_TB2P_SyncMode.ProfGenAbsolute;
	LRSLAVESYNCOUTPOS : LREAL := 0.0;
	LRSLAVESYNCINDIST : LREAL := 90.0;
	LRSLAVESYNCOUTDIST : LREAL := 90.0;
	LRSYNCVEL : LREAL := 100;
END_STRUCT
END_TYPE

(* ---- L_TS2P_SCPARSYNCHRONIZINGCAMMING.dut ---- *)
TYPE L_TS2P_SCPARSYNCHRONIZINGCAMMING :
STRUCT
	DWGEARINGNUMERATOR : DWORD := 1;
	DWGEARINGDENOMINATOR : DWORD := 1;
	LRSYNCACC : LREAL := 1000.0;
	LRSYNCDEC : LREAL := 1000.0;
	LRSYNCJERK : LREAL := 1000000.0;
	EALLOWEDDIRECTION : L_TB2P_AllowedDirection;
	XLIMITALLOWEDDIRECTION : BOOL := FALSE;
	LRTOLERANCEALLOWEDDIRECTION : LREAL := 5;
	LRSETOFFSETTRIMVEL : LREAL := 10.0;
	LRSETOFFSETTRIMACC : LREAL := 100.0;
	LRSETOFFSETTRIMDEC : LREAL := 100.0;
	LRSETOFFSETTRIMJERK : LREAL := 10000.0;
	XLOADOFFSET : BOOL;
	ETRIMMODE : L_TS2P_TrimMode := L_TS2P_TrimMode.position;
	LRTRIMDIST : LREAL := 1;
END_STRUCT
END_TYPE

(* ---- L_TS2P_SCSF_CROSSCUTTERBASE.dut ---- *)
TYPE L_TS2P_SCSF_CROSSCUTTERBASE :
STRUCT
END_STRUCT
END_TYPE

(* ---- L_TS2P_SCSF_CROSSCUTTERHIGH.dut ---- *)
TYPE L_TS2P_SCSF_CROSSCUTTERHIGH :
STRUCT
END_STRUCT
END_TYPE

(* ---- L_TS2P_SCSF_CROSSCUTTERSTATE.dut ---- *)
TYPE L_TS2P_SCSF_CROSSCUTTERSTATE :
STRUCT
END_STRUCT
END_TYPE

(* ---- L_TS2P_SCSF_ELECTRONICGEARBOXBASE.dut ---- *)
TYPE L_TS2P_SCSF_ELECTRONICGEARBOXBASE :
STRUCT
END_STRUCT
END_TYPE

(* ---- L_TS2P_SCSF_FLEXCAMHIGH.dut ---- *)
TYPE L_TS2P_SCSF_FLEXCAMHIGH :
STRUCT
END_STRUCT
END_TYPE

(* ---- L_TS2P_SCSF_FLEXCAMSTATE.dut ---- *)
TYPE L_TS2P_SCSF_FLEXCAMSTATE :
STRUCT
END_STRUCT
END_TYPE

(* ---- L_TS2P_SCSF_FLYINGSAWSTATE.dut ---- *)
TYPE L_TS2P_SCSF_FLYINGSAWSTATE :
STRUCT
END_STRUCT
END_TYPE

(* ---- L_TS2P_SCSF_SYNCANDCORRECTIONSTATE.dut ---- *)
TYPE L_TS2P_SCSF_SYNCANDCORRECTIONSTATE :
STRUCT
END_STRUCT
END_TYPE

(* ---- L_TS2P_SCSF_SYNCPOSBASE.dut ---- *)
TYPE L_TS2P_SCSF_SYNCPOSBASE :
STRUCT
END_STRUCT
END_TYPE

(* ---- L_TS2P_SCSF_TM_CROSSCUTTERBASE.dut ---- *)
TYPE L_TS2P_SCSF_TM_CROSSCUTTERBASE :
STRUCT
	MP_LWCHECKSUMENDOFPROFILE : LWORD;
	MP_LRSETMASTERPOS : LREAL;
	MP_LRCAMPROFILERPOSOUT : LREAL;
	MP_LRSETSLAVEPOSOUT : LREAL;
	MP_CAMPOINTSTART : ARRAY [0..3] OF L_MC2P_CamDataXYVA;
	MP_CAMPOINTCONTINUOUS : ARRAY [0..5] OF L_MC2P_CamDataXYVA;
	MP_CAMPOINTSTOP : ARRAY [0..3] OF L_MC2P_CamDataXYVA;
	MP_INUMOFPOINTSINCAM : INT;
	MP_BYSELECTCAM : BYTE;
	MP_BYSETTOOLNOOUT : BYTE;
	MP_BYSETAREAOUT : BYTE;
	MP_ECUTTINGPROCESSSTATE : L_TB2P_States;
	MP_LRYSTART : LREAL;
	MP_LRYPARK : LREAL;
	MP_LRYEND : LREAL;
	MP_LRXSTART : LREAL;
	MP_LRXENDSYNCPOS : LREAL;
	MP_LRXSTARTPARKPOS : LREAL;
	MP_LRXENDPARKPOS : LREAL;
	MP_LRXSTARTSYNCPOS : LREAL;
	MP_LRXEND : LREAL;
	MP_XXABSOLUTE : BOOL;
	MP_XSLAVEABSOLUTE : BOOL;
	MP_XENDOFPROFILE : BOOL;
	MP_XENDOFXCYCLE : BOOL;
	MP_XENABLEPOSITIONFOLLOWER : BOOL;
	MP_LROVERSPEED : LREAL;
	MP_LROFFSET : LREAL;
	MP_LROFFSETTRIM : LREAL;
	MP_LRSETXPOSOUT : LREAL;
	MP_LRSETXVELOUT : LREAL;
	MP_LRSETXACCOUT : LREAL;
	MP_LRSLAVEMAXVEL : LREAL;
	MP_LRSLAVEMAXACC : LREAL;
	MP_LRSETMOTORPRECTRLTRQOUT : LREAL;
	MP_XREGISTERCTRLACTIVE : BOOL;
END_STRUCT
END_TYPE

(* ---- L_TS2P_SCSF_TM_CROSSCUTTERHIGH.dut ---- *)
TYPE L_TS2P_SCSF_TM_CROSSCUTTERHIGH :
STRUCT
END_STRUCT
END_TYPE

(* ---- L_TS2P_SCSF_TM_CROSSCUTTERSTATE.dut ---- *)
TYPE L_TS2P_SCSF_TM_CROSSCUTTERSTATE :
STRUCT
	MP_XENABLETORQUEFOLLOWER : BOOL;
	MP_LRPRECTRLACCOUT : LREAL;
	MP_LRGEARBOXFACTOR : LREAL;
	MP_LRAXISTORQUE : LREAL;
	MP_LRINTEGRATORREGPOS : LREAL;
	MP_LRCORRREGPOS : LREAL;
	MP_LRMARKSENSORSETPOS : LREAL;
	MP_LRMARKACTTPPOS : LREAL;
	MP_XMARKRECEIVED : BOOL;
	MP_LRACTMARKERROR : LREAL;
	MP_LRACTMARKDIST : LREAL;
	MP_XCORRACTIVE : BOOL;
	MP_XCORRLIMITED : BOOL;
	MP_XMARKWINDOWOPEN : BOOL;
	MP_XMARKOUTOFWINDOW : BOOL;
	MP_XMARKNOTDETECTED : BOOL;
	MP_XGEARFACTORCORRLIMITED : BOOL;
	MP_LRSETCORRPOSOUT : LREAL;
	MP_LRSETCORRVELOUT : LREAL;
	MP_LRSETMASTERVEL : LREAL;
	MP_LRMARKSENSORSETPOSTOOL : LREAL;
	MP_LRMARKACTTPPOSTOOL : LREAL;
	MP_LRACTMARKERRORTOOL : LREAL;
	MP_XMARKRECEIVEDTOOL : BOOL;
	MP_XCORRACTIVETOOL : BOOL;
	MP_XCORRLIMITEDTOOL : BOOL;
	MP_XMARKWINDOWOPENTOOL : BOOL;
	MP_XMARKOUTOFWINDOWTOOL : BOOL;
	MP_XMARKNOTDETECTEDTOOL : BOOL;
	MP_XMARKWINDOWTEACHEDTOOL : BOOL;
END_STRUCT
END_TYPE

(* ---- L_TS2P_SCSF_TM_ELECTRONICGEARBOXBASE.dut ---- *)
TYPE L_TS2P_SCSF_TM_ELECTRONICGEARBOXBASE :
STRUCT
	MP_LRSETMASTERVEL : LREAL;
	MP_LRSETGEARBOXINVEL : LREAL;
	MP_LRSETGEARBOXOUTVEL : LREAL;
	MP_LRSETSLAVEVEL : LREAL;
	MP_LRVELOFFSET : LREAL;
	MP_LRPOSOFFSETTOTALPOS : LREAL;
	MP_LRPOSOFFSETTOTALVEL : LREAL;
	MP_LROFFSETTRIM : LREAL;
END_STRUCT
END_TYPE

(* ---- L_TS2P_SCSF_TM_FLEXCAM.dut ---- *)
TYPE L_TS2P_SCSF_TM_FLEXCAM :
STRUCT
	MP_LRSETMASTERPOS : LREAL;
	MP_LRSETMASTERVEL : LREAL;
	MP_LRSETCLUTCHPOSOUT : LREAL;
	MP_LRSETCLUTCHVELOUT : LREAL;
	MP_LRSETCLUTCHACCOUT : LREAL;
	MP_FINDCLUTCHXPOSACTIVE : BOOL;
	MP_FINDCLUTCHXPOSDONE : BOOL;
	MP_LWENDOFPROFILECHECKSUM : LWORD;
	MP_LRCONVERTMASTERTOXPOS : LREAL;
	MP_LRCAMPROFILERPOSOUT : LREAL;
	MP_LRSETXPOS : LREAL;
	MP_LRSETXVEL : LREAL;
	MP_LRSETXACC : LREAL;
	MP_LRSETYPOS : LREAL;
	MP_LRSETYVEL : LREAL;
	MP_LRSETYACC : LREAL;
	MP_LRCONVERTYTOSLAVEPOS : LREAL;
	MP_XENDOFPROFPOSITIVE : BOOL;
	MP_XENDOFPROFNEGATIVE : BOOL;
	MP_LRSLAVEMAXPOS : LREAL;
	MP_LRSLAVEMINPOS : LREAL;
	MP_LRSLAVEMAXVEL : LREAL;
	MP_LRSLAVEMAXACC : LREAL;
	MP_LRSETCAMPOSOUT : LREAL;
	MP_LRSETCAMVELOUT : LREAL;
	MP_LRSETCAMACCOUT : LREAL;
	MP_LRSETSYNCINPOSOUT : LREAL;
	MP_LRSETSYNCINVELOUT : LREAL;
	MP_LRSETSYNCINACCOUT : LREAL;
	MP_LRSETFOLLOWERPOS : LREAL;
	MP_LRSETFOLLOWERVEL : LREAL;
	MP_LRSETFOLLOWERACC : LREAL;
	MP_CAMTABLEACTIVE : MC_CAM_REF;
END_STRUCT
END_TYPE

(* ---- L_TS2P_SCSF_TM_FLEXCAMBASE.dut ---- *)
TYPE L_TS2P_SCSF_TM_FLEXCAMBASE :
STRUCT
	MP_LWENDOFPROFILECHECKSUM : LWORD;
	MP_LRSETMASTERPOS : LREAL;
	MP_LRSETSLAVEPOS : LREAL;
	MP_LRCONVERTMASTERTOXPOS : LREAL;
	MP_LRCAMPROFILERPOSOUT : LREAL;
	MP_LRCONVERTYTOSLAVEPOS : LREAL;
	MP_LRSETXPOS : LREAL;
	MP_LRSETXVEL : LREAL;
	MP_LRSETXACC : LREAL;
	MP_LRSETYPOS : LREAL;
	MP_LRSETYVEL : LREAL;
	MP_LRSETYACC : LREAL;
	MP_LRACTYPOS : LREAL;
	MP_LRACTYVEL : LREAL;
	MP_XENDOFPROFPOSITIVE : BOOL;
	MP_XENDOFPROFNEGATIVE : BOOL;
	MP_LRSLAVEMAXPOS : LREAL;
	MP_LRSLAVEMINPOS : LREAL;
	MP_LRSLAVEMAXVEL : LREAL;
	MP_LRSLAVEMAXACC : LREAL;
	MP_CAMTABLEACTIVE : MC_CAM_REF;
END_STRUCT
END_TYPE

(* ---- L_TS2P_SCSF_TM_FLEXCAMSTATE.dut ---- *)
TYPE L_TS2P_SCSF_TM_FLEXCAMSTATE :
STRUCT
END_STRUCT
END_TYPE

(* ---- L_TS2P_SCSF_TM_FLYINGSAWSTATE.dut ---- *)
TYPE L_TS2P_SCSF_TM_FLYINGSAWSTATE :
STRUCT
	MP_LRSETMASTERPOS : LREAL;
	MP_LRSETSLAVEPOS : LREAL;
	MP_LRTOTALCUTTINGLENGTH : LREAL;
	MP_XPOSSYNCHRONISED : BOOL;
	MP_LRCUTLENGTHPROCESSED : LREAL;
	MP_XMARKRECEIVED : BOOL;
	MP_WMARKINDEX : WORD;
	MP_XMARKSTACKEMPTY : BOOL;
	MP_XMARKSTACKFULL : BOOL;
	MP_MARKPOS : LREAL;
	MP_LRSTACKMARKPOS : LREAL;
	MP_XMASTERVELINWINDOW : BOOL;
	MP_XSLAVEPOSUPPERLIMIT : BOOL;
	MP_XSLAVEPOSLOWERLIMIT : BOOL;
END_STRUCT
END_TYPE

(* ---- L_TS2P_SCSF_TM_SYNCANDCORRECTIONSTATE.dut ---- *)
TYPE L_TS2P_SCSF_TM_SYNCANDCORRECTIONSTATE :
STRUCT
	MP_LRINTEGRATORREGPOS : LREAL;
	MP_LRCORRREGPOS : LREAL;
	MP_LRMARKSENSORSETPOS : LREAL;
	MP_LRMARKACTTPPOS : LREAL;
	MP_XMARKRECEIVED : BOOL;
	MP_LRACTMARKERROR : LREAL;
	MP_LRACTMARKDIST : LREAL;
	MP_XCORRACTIVE : BOOL;
	MP_XCORRLIMITED : BOOL;
	MP_XMARKWINDOWOPEN : BOOL;
	MP_XMARKOUTOFWINDOW : BOOL;
	MP_XMARKNOTDETECTED : BOOL;
	MP_LRGEARFACTORCORR : LREAL;
	MP_XGEARFACTORCORRLIMITED : BOOL;
	MP_LRSETCORRPOSOUT : LREAL;
	MP_LRSETCORRVELOUT : LREAL;
	MP_LRMARKSENSORSETPOSTOOL : LREAL;
	MP_LRMARKACTTPPOSTOOL : LREAL;
	MP_LRACTMARKERRORTOOL : LREAL;
	MP_XMARKRECEIVEDTOOL : BOOL;
	MP_XCORRACTIVETOOL : BOOL;
	MP_XCORRLIMITEDTOOL : BOOL;
	MP_XMARKWINDOWOPENTOOL : BOOL;
	MP_XMARKOUTOFWINDOWTOOL : BOOL;
	MP_XMARKNOTDETECTEDTOOL : BOOL;
	MP_XMARKWINDOWTEACHEDTOOL : BOOL;
END_STRUCT
END_TYPE

(* ---- L_TS2P_SCSF_TM_SYNCPOSBASE.dut ---- *)
TYPE L_TS2P_SCSF_TM_SYNCPOSBASE :
STRUCT
	MP_LRSETMASTERPOS : LREAL;
	MP_LRSETMASTERVEL : LREAL;
	MP_LRSETGEARBOXPOSIN : LREAL;
	MP_LRSETGEARBOXVELIN : LREAL;
	MP_LRSETGEARBOXPOSOUT : LREAL;
	MP_LRSETGEARBOXVELOUT : LREAL;
	MP_LRSETCLUTCHPOSIN : LREAL;
	MP_LROFFSET : LREAL;
	MP_LROFFSETTRIM : LREAL;
	MP_LROFFSETTOTALVEL : LREAL;
	MP_LROFFSETSYNCPOS : LREAL;
END_STRUCT
END_TYPE

(* ---- L_TS2P_SOURCEFORCORRWINDOW.dut ---- *)
TYPE L_TS2P_SOURCEFORCORRWINDOW :
(
	CORRECTEDMASTERPOS := 1,
	SLAVE := 2
);
END_TYPE

(* ---- L_TS2P_SYNCANDCORRECTIONSTATEIN.dut ---- *)
TYPE L_TS2P_SYNCANDCORRECTIONSTATEIN :
STRUCT
	SCTPRECDATA_MARKSENSOR : L_MC1P_TpReceiveData;
	SCTPRECDATA_TOOLSENSOR : L_MC1P_TpReceiveData;
	XTEACHMARKWINDOW : BOOL;
	XTEACHMARKWINDOWTOOL : BOOL;
	XGEARFACTORCORR : BOOL;
	XGEARFACTORCORRHOLD : BOOL;
END_STRUCT
END_TYPE

(* ---- L_TS2P_SYNCANDCORRECTIONSTATEOUT.dut ---- *)
TYPE L_TS2P_SYNCANDCORRECTIONSTATEOUT :
STRUCT
	LRSETMARKCORROUT : LREAL;
	XMARKWINDOWTEACHED : BOOL;
	LRGEARFACTORCORR : LREAL;
	LRSETTOOLCORROUT : LREAL;
	XMARKWINDOWTEACHEDTOOL : BOOL;
END_STRUCT
END_TYPE

(* ---- L_TS2P_SYNCDIRECTION.dut ---- *)
TYPE L_TS2P_SYNCDIRECTION :
(
	POSITIVEDIRECTION := 1,
	NEGATIVEDIRECTION := 2,
	SHORTESTWAY := 3
);
END_TYPE

(* ---- L_TS2P_SYNCINMODE.dut ---- *)
TYPE L_TS2P_SYNCINMODE :
(
	PROFGENABSOLUTE := 0,
	PROFGENRELATIVE := 1
);
END_TYPE

(* ---- L_TS2P_SYNCMODECROSSCUTTER.dut ---- *)
TYPE L_TS2P_SYNCMODECROSSCUTTER :
(
	CAM_IN := 0,
	POSITIONING := 1
);
END_TYPE

(* ---- L_TS2P_SYNCMODEFLEXCAM.dut ---- *)
TYPE L_TS2P_SYNCMODEFLEXCAM :
(
	PROFGENABSOLUTE := 0,
	CAMABSOLUTE := 4,
	INSTANTABSOLUTE := 10,
	INSTANTRELATIVE := 11
);
END_TYPE

(* ---- L_TS2P_SYNCPOSBASEIN.dut ---- *)
TYPE L_TS2P_SYNCPOSBASEIN :
STRUCT
	MASTERVALUES : L_MC1P_IAXIS_REF_MASTERVALUES;
	XSYNCIN : BOOL;
	XSYNCPOSRESTORE : BOOL;
	LRSETBASEVEL : LREAL;
	LRSETOFFSETPOS : LREAL;
	XTRIMPOS : BOOL;
	XTRIMNEG : BOOL;
	XTRIMRESET : BOOL;
END_STRUCT
END_TYPE

(* ---- L_TS2P_SYNCPOSBASEOUT.dut ---- *)
TYPE L_TS2P_SYNCPOSBASEOUT :
STRUCT
	XSYNCHRONISED : BOOL;
	XACCDECSYNC : BOOL;
	XOFFSETTRIMACTIVE : BOOL;
	XBASEVELOCITYACTIVE : BOOL;
	LROFFSETTOTAL : LREAL;
END_STRUCT
END_TYPE

(* ---- L_TS2P_TRIMMODE.dut ---- *)
TYPE L_TS2P_TRIMMODE :
(
	VELOCITY := 0,
	POSITION := 1
);
END_TYPE

(* ---- L_TS2P_XYBUFFERDATA.dut ---- *)
TYPE L_TS2P_XYBUFFERDATA :
STRUCT
	LRBUFFERPOSITIONPOS : LREAL;
	LRBUFFERPOSITIONNEG : LREAL;
	LRBUFFERVELPOS : LREAL;
	LRBUFFERVELNEG : LREAL;
END_STRUCT
END_TYPE

(* ---- L_TS2P_XYLIMITS.dut ---- *)
TYPE L_TS2P_XYLIMITS :
STRUCT
	LRVELOCITY : LREAL;
	LRACCELERATION : LREAL;
	LRDECELERATION : LREAL;
END_STRUCT
END_TYPE

(* ---- L_TS2P_INTERNAL.gvl ---- *)
VAR_GLOBAL
	CDIENUMSTARTVALUE : DINT := 22000;
END_VAR

(* ---- L_TS2M_ITFFLYINGSAWSTATEFMDATA.itf ---- *)
INTERFACE L_TS2M_ITFFLYINGSAWSTATEFMDATA
END_INTERFACE

(* ---- L_TS2M_ITFFLYINGSAWSTATETMDATA.itf ---- *)
INTERFACE L_TS2M_ITFFLYINGSAWSTATETMDATA
END_INTERFACE

METHOD MOVETOPARKPOS : BOOL
VAR_INPUT
	XEXECUTEMOVETOPARKPOS : BOOL;
	LRPARKPOSITION : LREAL := 180;
	EPOSITIONINGDIRECTION : MC_DIRECTION := MC_DIRECTION.mcPositiveDirection;
	LRPOSITIONINGVEL : LREAL := 10;
	LRPOSITIONINGACC : LREAL := 100;
	LRPOSITIONINGDEC : LREAL := 100;
	LRJERK : LREAL := 0;
END_VAR
VAR_OUTPUT
	XBUSY : BOOL;
	XDONE : BOOL;
	XCOMMANDABORTED : BOOL;
END_VAR
VAR_IN_OUT
	AXIS : AXIS_REF;
END_VAR
END_METHOD

(* ---- L_TS2P_ICONNECTORFLEXCAM.itf ---- *)
INTERFACE L_TS2P_ICONNECTORFLEXCAM
END_INTERFACE

(* ---- L_TS2P_ICONNECTORFLYINGSAW.itf ---- *)
INTERFACE L_TS2P_ICONNECTORFLYINGSAW
END_INTERFACE

(* ---- L_TS2P_ICONNECTORSYNCANDCORRECTION.itf ---- *)
INTERFACE L_TS2P_ICONNECTORSYNCANDCORRECTION
END_INTERFACE

(* ---- L_TS2P_ICONNECTORSYNCPOS.itf ---- *)
INTERFACE L_TS2P_ICONNECTORSYNCPOS
END_INTERFACE

(* ---- L_TS2P_IFLEXCAM.itf ---- *)
INTERFACE L_TS2P_IFLEXCAM
END_INTERFACE

METHOD CAM
VAR_INPUT
	ITFTECHMODULE : L_TS2P_IFlexCam;
	XENABLE : BOOL;
	XSYNCCAM : BOOL;
	SCCAMTABLE : MC_CAM_REF;
	LRCYCMASTERPOS : LREAL;
	LRCYCMASTERVEL : LREAL;
	LRCYCMASTERACC : LREAL;
	LRSLAVEPOS : LREAL;
	LRSLAVEVEL : LREAL;
	LRSLAVEACC : LREAL;
	EOFFSETMODEMASTER : L_TS2P_OffsetMode := L_TS2P_OffsetMode.x_zero;
	ESCALINGMODEMASTER : L_TS2P_ScalingMode := L_TS2P_ScalingMode.x_zero;
	EOFFSETMODESLAVE : L_TS2P_OffsetMode := L_TS2P_OffsetMode.x_zero;
	ESCALINGMODESLAVE : L_TS2P_ScalingMode := L_TS2P_ScalingMode.x_zero;
	LRSETOFFSETMASTER : LREAL;
	LRSETOFFSETSLAVE : LREAL;
	LRSETSCALINGMASTER : LREAL;
	LRSETSCALINGSLAVE : LREAL;
	LRPROFGENMASTERVEL : LREAL;
	LRPROFGENMASTERACC : LREAL;
	LRPROFGENMASTERDEC : LREAL;
	LRPROFGENMASTERJERK : LREAL;
	LRPROFGENSLAVEVEL : LREAL;
	LRPROFGENSLAVEACC : LREAL;
	LRPROFGENSLAVEDEC : LREAL;
	LRPROFGENSLAVEJERK : LREAL;
	XPERIODIC : BOOL;
	XCAMCHANGEINSTANT : BOOL;
	XMASTERABSOLUTE : BOOL;
	XSLAVEABSOLUTE : BOOL;
END_VAR
VAR_OUTPUT
	XERROR : BOOL;
	EERRORID : L_IE1P.L_IE1P_Error;
	LRSETPOSOUT : LREAL;
	LRSETVELOUT : LREAL;
	LRSETACCOUT : LREAL;
	LRSETXPOSOUT : LREAL;
	LRSETXVELOUT : LREAL;
	LRSETXACCOUT : LREAL;
	LRSETYPOSOUT : LREAL;
	LRSETYVELOUT : LREAL;
	LRSETYACCOUT : LREAL;
	XENDOFPROFILE : BOOL;
	LRSETOFFSETMASTEROUT : LREAL;
	LRSETOFFSETSLAVEOUT : LREAL;
	LRCONVERTMASTERTOXPOS : LREAL;
	LRCAMPROFILERPOSOUT : LREAL;
	LRCONVERTYTOSLAVEPOS : LREAL;
	XDONE : BOOL;
	XBUSY : BOOL;
END_VAR
END_METHOD

METHOD CAMSEQUENCER
VAR_INPUT
	ITFTECHMODULE : L_TS2P_IFlexCam;
	XENABLE : BOOL;
	XCAMSEQUENCER : BOOL;
	XENDOFPROFILEIN : BOOL;
	CAMTABLE1 : MC_CAM_REF;
	CAMTABLE2 : MC_CAM_REF;
	CAMTABLE3 : MC_CAM_REF;
	CAMTABLE4 : MC_CAM_REF;
	XCAMCHANGEINSTANT : BOOL;
	XLOADCAMTABLE : BOOL;
	WSETCAMTABLE : WORD;
	EMODE : L_TS2P_CamSequenceMode := L_TS2P_CamSequenceMode.CyclicCam1;
END_VAR
VAR_OUTPUT
	XERROR : BOOL;
	EERRORID : L_IE1P_Error;
	CAMTABLEOUT : MC_CAM_REF;
	XCAMTABLEVALID : BOOL;
END_VAR
END_METHOD

METHOD CLUTCH
VAR_INPUT
	ITFTECHMODULE : L_TS2P_IFlexCam;
	XENABLE : BOOL;
	XCLUTCHCLOSE : BOOL;
	ECLUTCHINMODE : L_TS2P_ClutchInMode;
	ECLUTCHOUTMODE : L_TS2P_ClutchOutMode;
	EALLOWEDDIRECTION : L_TB2P_AllowedDirection;
	LRCLUTCHINDIST : LREAL;
	LRCLUTCHOUTDIST : LREAL;
	LRCLUTCHOUTPOSITION : LREAL;
	LRCYCLICMASTERPOS : LREAL;
	LRCYCLICMASTERVEL : LREAL;
	LRCYCLICMASTERACC : LREAL;
	LRCYCLICAXISPOS : LREAL;
	LRCYCLICAXISVEL : LREAL;
	LRCYCLICAXISACC : LREAL;
	ETRAVERSINGRANGE : L_MC1P_TraversingRange;
	LRCYCLELENGTH : LREAL;
END_VAR
VAR_OUTPUT
	XERROR : BOOL;
	EERRORID : L_IE1P.L_IE1P_Error;
	XBUSY : BOOL;
	XDONE : BOOL;
	XSYNCHRONISED : BOOL;
	XACCDECSYNC : BOOL;
	LRSETPOSOUT : LREAL;
	LRSETVELOUT : LREAL;
	LRSETACCOUT : LREAL;
END_VAR
END_METHOD

METHOD HALT : BOOL
VAR_INPUT
	ITFTECHMODULE : L_TS2P_IFlexCam;
	XEXECUTE : BOOL;
	LRDEC : LREAL := 100;
	LRJERK : LREAL := 0;
END_VAR
VAR_OUTPUT
	XBUSY : BOOL;
	XDONE : BOOL;
	XCOMMANDABORTED : BOOL;
END_VAR
VAR_IN_OUT
	AXIS : AXIS_REF;
END_VAR
END_METHOD

METHOD MOVETOPARKPOS : BOOL
VAR_INPUT
	ITFTECHMODULE : L_TS2P_IFlexCam;
	XEXECUTEMOVETOPARKPOS : BOOL;
	EMOVETOPARKPOSMODE : L_TS2P_CamStopMode;
	LRPARKPOSITION : LREAL := 180;
	EPOSITIONINGDIRECTION : L_TS2P_SyncDirection := L_TS2P_SyncDirection.PositiveDirection;
	LRPOSITIONINGVEL : LREAL := 10;
	LRPOSITIONINGACC : LREAL := 100;
	LRPOSITIONINGDEC : LREAL := 100;
	LRJERK : LREAL := 0;
END_VAR
VAR_OUTPUT
	XBUSY : BOOL;
	XDONE : BOOL;
	XCOMMANDABORTED : BOOL;
END_VAR
VAR_IN_OUT
	AXIS : AXIS_REF;
END_VAR
END_METHOD

METHOD POSITIONFOLLOWER
VAR_INPUT
	ITFTECHMODULE : L_TS2P_IFlexCam;
	XENABLE : BOOL;
	LRPOSITION : LREAL;
	LRVELOCITY : LREAL;
	LRACCELERATION : LREAL;
	ESETVALUEMODE : L_MC1P_SetValueMode;
END_VAR
VAR_OUTPUT
	XERROR : BOOL;
	EERRORID : L_IE1P.L_IE1P_Error;
	XBUSY : BOOL;
END_VAR
END_METHOD

METHOD SYNCIN
VAR_INPUT
	ITFTECHMODULE : L_TS2P_IFlexCam;
	XENABLE : BOOL;
	XSYNCIN : BOOL;
	XSYNCPOSRESTORE : BOOL;
	ESYNCMODE : L_TS2P_SyncInMode;
	ESYNCDIRECTION : L_TS2P_SyncDirection;
	LRSYNCVEL : LREAL;
	LRSYNCACC : LREAL;
	LRSYNCDEC : LREAL;
	LRSYNCJERK : LREAL;
	LRPARKPOSITION : LREAL;
	LRCYCLICMASTERPOS : LREAL;
	LRCYCLICMASTERVEL : LREAL;
	LRCYCLICMASTERACC : LREAL;
	LRCYCLICAXISPOS : LREAL;
	LRCYCLICAXISVEL : LREAL;
	LRCYCLICAXISACC : LREAL;
END_VAR
VAR_OUTPUT
	XERROR : BOOL;
	EERRORID : L_IE1P.L_IE1P_Error;
	XBUSY : BOOL;
	XDONE : BOOL;
	XSYNCHRONISED : BOOL;
	XACCDECSYNC : BOOL;
	LRSETPOSOUT : LREAL;
	LRSETVELOUT : LREAL;
	LRSETACCOUT : LREAL;
	LROFFSETSYNCPOS : LREAL;
END_VAR
VAR_IN_OUT
	AXIS : AXIS_REF;
END_VAR
END_METHOD

(* ---- L_TS2P_IFLYINGSAWPROCESSING.itf ---- *)
INTERFACE L_TS2P_IFLYINGSAWPROCESSING
END_INTERFACE

METHOD CLUTCH
VAR_INPUT
	ITFTECHMODULE : L_TS2P_IFlyingSawProcessing;
	XENABLE : BOOL;
	XSYNCVEL : BOOL := FALSE;
	XSYNCPOS : BOOL;
	XSYNCOUTINSTANT : BOOL;
	LRSYNCVEL : LREAL := 10;
	LRSYNCACC : LREAL := 100;
	LRSYNCDEC : LREAL := 100;
	LRSYNCJERK : LREAL := 10000;
	LRCYCMASTERPOS : LREAL;
	LRCYCMASTERVEL : LREAL;
	LRCYCMASTERACC : LREAL;
	LRSETSLAVEPOS : LREAL;
	LRSETSLAVEVEL : LREAL;
	LRSETSLAVEACC : LREAL;
END_VAR
VAR_OUTPUT
	EERRORID : L_IE1P_Error;
	XERROR : BOOL;
	XBUSY : BOOL;
	XDONE : BOOL;
	XACCDECSYNC : BOOL;
	XVELSYNCHRONISED : BOOL;
	XPOSSYNCHRONISED : BOOL;
	LRSETSLAVEPOSOUT : LREAL;
	LRSETSLAVEVELOUT : LREAL;
	LRSETSLAVEACCOUT : LREAL;
	XPROFILERESETTIMEVALID : BOOL;
	LRPROFILERESETTIME : LREAL;
END_VAR
END_METHOD

METHOD EXECUTEGAP
VAR_INPUT
	ITFTECHMODULE : L_TS2P_IFlyingSawProcessing;
	XENABLE : BOOL;
	LRSYNCVEL : LREAL := 10;
	LRSYNCACC : LREAL := 100;
	LRSYNCDEC : LREAL := 100;
	LRSYNCJERK : LREAL := 10000;
	XEXECUTEGAP : BOOL;
	XAUXEXECUTEGAP : BOOL := FALSE;
	LRCYCMASTERPOS : LREAL;
	LRCYCMASTERVEL : LREAL;
	LRCYCMASTERACC : LREAL;
	LRSETSLAVEPOS : LREAL;
	LRSETSLAVEVEL : LREAL;
	LRSETSLAVEACC : LREAL;
END_VAR
VAR_OUTPUT
	EERRORID : L_IE1P_Error;
	XERROR : BOOL;
	XBUSY : BOOL;
	XDONE : BOOL;
	XACCDECSYNC : BOOL;
	XVELSYNCHRONISED : BOOL;
	XPOSSYNCHRONISED : BOOL;
	LRSETSLAVEPOSOUT : LREAL;
	LRSETSLAVEVELOUT : LREAL;
	LRSETSLAVEACCOUT : LREAL;
	XPROFILERESETTIMEVALID : BOOL;
	LRPROFILERESETTIME : LREAL;
END_VAR
END_METHOD

METHOD MARKSTACK_GETMARK
VAR_INPUT
	ITFTECHMODULE : L_TS2P_IFlyingSawProcessing;
	XENABLE : BOOL;
	XGETMARK : BOOL;
	XRESETGETMARK : BOOL;
	XRESETMARKSTACK : BOOL;
	LRCYCSETPOS : LREAL;
	LRCYCSETVEL : LREAL;
END_VAR
VAR_OUTPUT
	XMARKSTACKFULL : BOOL;
	XMARKSTACKEMPTY : BOOL;
	WMARKSINSTACK : WORD;
	XMARKVALID : BOOL;
	LRMARKPOSOUT : LREAL;
END_VAR
END_METHOD

METHOD MARKSTACK_SETMARK
VAR_INPUT
	ITFTECHMODULE : L_TS2P_IFlyingSawProcessing;
	XENABLE : BOOL;
	XSETMARK : BOOL;
	LRMARKPOS : LREAL;
	XRESETMARKSTACK : BOOL;
	LRCYCSETPOS : LREAL;
	LRCYCSETVEL : LREAL;
END_VAR
VAR_OUTPUT
	XMARKSTACKFULL : BOOL;
	XMARKSTACKEMPTY : BOOL;
	WMARKSINSTACK : WORD;
	XNEWMARKRECEIVED : BOOL;
END_VAR
END_METHOD

METHOD POSITIONING
VAR_INPUT
	ITFTECHMODULE : L_TS2P_IFlyingSawProcessing;
	XENABLE : BOOL;
	XMOVETOTARGETPOS : BOOL;
	LRTARGETPOS : LREAL;
	LRPOSITIONINGVEL : LREAL;
	LRPOSITIONINGACC : LREAL;
	LRPOSITIONINGDEC : LREAL;
	LRPOSITIONINGJERK : LREAL;
	LRSETSLAVEPOS : LREAL;
	LRSETSLAVEVEL : LREAL;
	LRSETSLAVEACC : LREAL;
	LRCORRECTTIMEBASE : LREAL := 0;
	LROVERRIDE : LREAL := 1.0;
END_VAR
VAR_OUTPUT
	EERRORID : L_IE1P_Error;
	XERROR : BOOL;
	XBUSY : BOOL;
	XDONE : BOOL;
	XPOSITIONING : BOOL;
	XINPOSITION : BOOL;
	LRSETSLAVEPOSOUT : LREAL;
	LRSETSLAVEVELOUT : LREAL;
	LRSETSLAVEACCOUT : LREAL;
	XPROFILERESETTIMEVALID : BOOL;
	LRPROFILERESETTIME : LREAL;
END_VAR
END_METHOD

(* ---- L_TS2P_ISIGNALFLOW.itf ---- *)
INTERFACE L_TS2P_ISIGNALFLOW
END_INTERFACE

METHOD GET_PSF : POINTER TO L_TS2P_scSF_TM_SyncPosBase
END_METHOD

(* ---- L_TS2P_ISIGNALFLOWFLEXCAM.itf ---- *)
INTERFACE L_TS2P_ISIGNALFLOWFLEXCAM
END_INTERFACE

METHOD GET_PSF : POINTER TO L_TS2P_scSF_TM_SyncPosBase
END_METHOD

(* ---- L_TS2P_ISIGNALFLOWSC.itf ---- *)
INTERFACE L_TS2P_ISIGNALFLOWSC
END_INTERFACE

METHOD GET_PSF : POINTER TO L_TS2P_scSF_TM_SyncAndCorrectionState
END_METHOD

(* ---- L_TS2P_ISTRUCTPROVIDERFLEXCAMHIGH.itf ---- *)
INTERFACE L_TS2P_ISTRUCTPROVIDERFLEXCAMHIGH
END_INTERFACE

METHOD GET_PDATA : POINTER TO L_TS2P_scData_TM_FlexCam
END_METHOD

METHOD GET_PDATASP : POINTER TO L_TS2P_scData_TM_FlexCam
END_METHOD

(* ---- L_TS2P_ISTRUCTPROVIDERFLYINGSAW.itf ---- *)
INTERFACE L_TS2P_ISTRUCTPROVIDERFLYINGSAW
END_INTERFACE

METHOD GET_PDATA : POINTER TO L_TS2M_scData_FlyingSawState
END_METHOD

METHOD GET_PFMDATA : POINTER TO L_TS2M_scData_FM_FlyingSaw
END_METHOD

(* ---- L_TS2P_ISTRUCTPROVIDERSYNCANDCORRECTION.itf ---- *)
INTERFACE L_TS2P_ISTRUCTPROVIDERSYNCANDCORRECTION
END_INTERFACE

METHOD GET_PDATA : POINTER TO L_TS2P_scData_TM_SyncAndCorrectionState
END_METHOD

METHOD GET_PDATASP : POINTER TO L_TS2P_scData_TM_SyncPosBase
END_METHOD

(* ---- L_TS2P_ISTRUCTPROVIDERSYNCPOS.itf ---- *)
INTERFACE L_TS2P_ISTRUCTPROVIDERSYNCPOS
END_INTERFACE

METHOD GET_PDATA : POINTER TO L_TS2P_scData_TM_SyncPosBase
END_METHOD

(* ---- L_TS2P_ISYNCANDCORRECTIONSTATE.itf ---- *)
INTERFACE L_TS2P_ISYNCANDCORRECTIONSTATE
END_INTERFACE

(* ---- L_TS2P_ISYNCPOSBASE.itf ---- *)
INTERFACE L_TS2P_ISYNCPOSBASE
END_INTERFACE

METHOD ADDOFFSET
VAR_INPUT
	ITFTECHMODULE : L_TS2P_ISyncPosBase;
	LRSETPOS : LREAL;
	LRSETVEL : LREAL;
	LRSETOFFSET : LREAL;
	LRSETOFFSETVEL : LREAL;
	ETRAVERSINGRANGE : L_MC1P.L_MC1P_TraversingRange;
	LRCYCLELENGTH : LREAL;
END_VAR
VAR_OUTPUT
	XERROR : BOOL;
	EERRORID : L_IE1P.L_IE1P_Error;
	LRSETPOSOUT : LREAL;
	LRSETVELOUT : LREAL;
END_VAR
END_METHOD

METHOD CLUTCH
VAR_INPUT
	ITFTECHMODULE : L_TS2P_ISyncPosBase;
	XENABLE : BOOL;
	XSYNCIN : BOOL;
	LRSETBASEVELOCITY : LREAL;
	ESYNCMODE : L_TB2P_SyncMode;
	EALLOWEDDIRECTION : L_TB2P_AllowedDirection;
	LRSYNCVEL : LREAL;
	LRSYNCACC : LREAL;
	LRSYNCDEC : LREAL;
	LRSYNCJERK : LREAL;
	LRSYNCINDIST : LREAL;
	LRSYNCOUTDIST : LREAL;
	LRSYNCOUTPOS : LREAL;
	XLOADCLUTCHOFFSET : BOOL;
	LRLOADCLUTCHOFFSET : LREAL;
	LRCYCLICMASTERPOS : LREAL;
	LRCYCLICMASTERVEL : LREAL;
	ETRAVERSINGRANGEMASTER : L_MC1P_TraversingRange;
	LRCYCLELENGTHMASTER : LREAL;
	LRCYCLICAXISPOS : LREAL;
	LRCYCLICAXISVEL : LREAL;
	LRCYCLICAXISACC : LREAL;
	ETRAVERSINGRANGEAXIS : L_MC1P_TraversingRange;
	LRCYCLELENGTHAXIS : LREAL;
END_VAR
VAR_OUTPUT
	XERROR : BOOL;
	EERRORID : L_IE1P.L_IE1P_Error;
	XBUSY : BOOL;
	XDONE : BOOL;
	XSYNCHRONISED : BOOL;
	XACCDECSYNC : BOOL;
	XINBASEVELOCITY : BOOL;
	LRSETPOSOUT : LREAL;
	LRSETVELOUT : LREAL;
	LRSETACCOUT : LREAL;
	LRCLUTCHOFFSETOUT : LREAL;
END_VAR
END_METHOD

METHOD GEARBOX
VAR_INPUT
	ITFTECHMODULE : L_TS2P_ISyncPosBase;
	XENABLE : BOOL;
	LRSETPOSX : LREAL;
	LRSETVELX : LREAL;
	DWNUMERATOR : DWORD;
	DWDENOMINATOR : DWORD;
	LRCYCLELENGTHX : LREAL;
	LRCYCLELENGTHY : LREAL;
	ETRAVERSINGRANGEX : L_MC1P.L_MC1P_TraversingRange;
	ETRAVERSINGRANGEY : L_MC1P.L_MC1P_TraversingRange;
	XLOADGEARBOXPOS : BOOL;
	LRLOADGEARBOXPOS : LREAL;
END_VAR
VAR_OUTPUT
	XERROR : BOOL;
	EERRORID : L_IE1P.L_IE1P_Error;
	LRSETPOSOUT : LREAL;
	LRSETVELOUT : LREAL;
END_VAR
END_METHOD

METHOD OFFSETANDTRIM
VAR_INPUT
	ITFTECHMODULE : L_TS2P_ISyncPosBase;
	XENABLE : BOOL;
	LRSETOFFSET : LREAL;
	XTRIMPOS : BOOL;
	XTRIMNEG : BOOL;
	LRSETTRIMDISTANCE : LREAL;
	ETRIMMODE : L_TS2P_TrimMode;
	XLOADOFFSET : BOOL;
	XRESETTRIMOFFSET : BOOL;
	LRSETVEL : LREAL;
	LRSETACC : LREAL;
	LRSETDEC : LREAL;
	LRSETJERK : LREAL;
	WACTDIRECTION : WORD;
	EALLOWEDDIRECTION : L_TB2P.L_TB2P_AllowedDirection;
	LRCYCMASTERPOS : LREAL;
	LRCYCMASTERVEL : LREAL;
	LRCYCMASTERACC : LREAL;
END_VAR
VAR_OUTPUT
	XERROR : BOOL;
	EERRORID : L_IE1P.L_IE1P_Error;
	XBUSY : BOOL;
	XDONE : BOOL;
	LRSETOFFSETOUTTOTAL : LREAL;
	LRSETOFFSETOUTTOTALVEL : LREAL;
	LRSETOFFSETOUT : LREAL;
	LRSETOFFSETOUTTRIM : LREAL;
END_VAR
END_METHOD

(* ---- GETBOOLEANPROPERTY.pou ---- *)
FUNCTION GETBOOLEANPROPERTY : BOOL
VAR_INPUT
	STKEY : WSTRING;
END_VAR
END_FUNCTION

(* ---- GETCOMPANY.pou ---- *)
FUNCTION GETCOMPANY : WSTRING
END_FUNCTION

(* ---- GETNUMBERPROPERTY.pou ---- *)
FUNCTION GETNUMBERPROPERTY : DINT
VAR_INPUT
	STKEY : WSTRING;
END_VAR
END_FUNCTION

(* ---- GETTEXTPROPERTY.pou ---- *)
FUNCTION GETTEXTPROPERTY : WSTRING
VAR_INPUT
	STKEY : WSTRING;
END_VAR
END_FUNCTION

(* ---- GETTEXTPROPERTY2.pou ---- *)
FUNCTION GETTEXTPROPERTY2 : POINTER TO WSTRING
VAR_INPUT
	STKEY : WSTRING;
END_VAR
END_FUNCTION

(* ---- GETTITLE.pou ---- *)
FUNCTION GETTITLE : WSTRING
END_FUNCTION

(* ---- GETVERSION.pou ---- *)
FUNCTION GETVERSION : VERSION
END_FUNCTION

(* ---- GETVERSIONPROPERTY.pou ---- *)
FUNCTION GETVERSIONPROPERTY : VERSION
VAR_INPUT
	STKEY : WSTRING;
END_VAR
END_FUNCTION

(* ---- L_MB1P_CONVERTPOSTOMODULOPOS.pou ---- *)
FUNCTION L_MB1P_CONVERTPOSTOMODULOPOS : LREAL
VAR_INPUT
	LRPOS : LREAL;
	LRPERIOD : LREAL;
END_VAR
VAR_OUTPUT
	DIREVCOUNTER : DINT;
END_VAR
END_FUNCTION

(* ---- L_MB1P_CONVERTPOSTOMODULOPOSEXTENDED.pou ---- *)
FUNCTION L_MB1P_CONVERTPOSTOMODULOPOSEXTENDED : LREAL
VAR_INPUT
	LRPOS : LREAL;
	LRPERIOD : LREAL;
END_VAR
VAR_OUTPUT
	DIREVCOUNTER : DINT;
END_VAR
END_FUNCTION

(* ---- L_MB1P_CONVERTPOSTOMODULOPOSFMOD.pou ---- *)
FUNCTION L_MB1P_CONVERTPOSTOMODULOPOSFMOD : LREAL
VAR_INPUT
	LRPOS : LREAL;
	LRPERIOD : LREAL;
END_VAR
END_FUNCTION

(* ---- L_MB1P_HLPCALCKOEFPOLY5THORD.pou ---- *)
FUNCTION L_MB1P_HLPCALCKOEFPOLY5THORD : ARRAY [0..5] OF LREAL
VAR_INPUT
	LRYPOSSTART : LREAL;
	LRYVELSTART : LREAL;
	LRYACCSTART : LREAL;
	LRYPOSEND : LREAL;
	LRYVELEND : LREAL;
	LRYACCEND : LREAL;
END_VAR
VAR_OUTPUT
	ALRKOEF : ARRAY [0..5] OF LREAL;
END_VAR
END_FUNCTION

(* ---- L_MB1P_HLPCALCYOFPOLY5THORDBASE.pou ---- *)
FUNCTION L_MB1P_HLPCALCYOFPOLY5THORDBASE : LREAL
VAR_OUTPUT
	LRYPOSSCALED : LREAL;
END_VAR
VAR_IN_OUT
	LRXPOSSCALED : LREAL;
	ALRKOEF : ARRAY [0..5] OF LREAL;
END_VAR
END_FUNCTION

(* ---- L_MB1P_HLPCALCYOFPOLY5THORDSTATE.pou ---- *)
FUNCTION L_MB1P_HLPCALCYOFPOLY5THORDSTATE : LREAL
VAR_INPUT
	LRXPOSSTART : LREAL;
	LRXPOSEND : LREAL := 1;
	LRSETXPOS : LREAL;
	ALRKOEF : ARRAY [0..5] OF LREAL;
END_VAR
VAR_OUTPUT
	LRYPOSSCALED : LREAL;
END_VAR
END_FUNCTION

(* ---- L_MB1P_HLPDELTAVELTIMEEXTENDED.pou ---- *)
FUNCTION L_MB1P_HLPDELTAVELTIMEEXTENDED : BOOL
VAR_INPUT
	LRVELSTART : LREAL;
	LRACCSTART : LREAL;
	LRMAXACC : LREAL;
	LRMAXJERK : LREAL;
END_VAR
VAR_OUTPUT
	LRTIME : LREAL;
	LRDIST : LREAL;
END_VAR
END_FUNCTION

(* ---- L_MB1P_HLPDELTAVELTIMESTATE.pou ---- *)
FUNCTION L_MB1P_HLPDELTAVELTIMESTATE : BOOL
VAR_INPUT
	LRVELSTART : LREAL;
	LRACCSTART : LREAL;
	LRVELTARGET : LREAL;
	LRACCTARGET : LREAL;
	LRMAXACC : LREAL;
	LRMAXDEC : LREAL;
	LRMAXJERK : LREAL;
END_VAR
VAR_OUTPUT
	LRTIME : LREAL;
	LRDIST : LREAL;
END_VAR
END_FUNCTION

(* ---- L_MB1P_HLPDELTAVELTIMETOCONTANTVEL.pou ---- *)
FUNCTION L_MB1P_HLPDELTAVELTIMETOCONTANTVEL : BOOL
VAR_INPUT
	LRACCSTART : LREAL;
	LRMAXJERK : LREAL;
	WMODE : WORD;
END_VAR
VAR_OUTPUT
	LRVEL : LREAL;
	LRTIME : LREAL;
	LRDIST : LREAL;
END_VAR
END_FUNCTION

(* ---- L_MB1P_HLPRESTTIMEFORDISTANCE.pou ---- *)
FUNCTION L_MB1P_HLPRESTTIMEFORDISTANCE : BOOL
VAR_OUTPUT
	LRTIME : LREAL;
END_VAR
VAR_IN_OUT
	LRVELSTART : LREAL;
	LRACCSTART : LREAL;
	LRDIST : LREAL;
END_VAR
END_FUNCTION

(* ---- L_MB1P_MODULOCYCLE.pou ---- *)
FUNCTION L_MB1P_MODULOCYCLE : LREAL
VAR_INPUT
	LRPOSIN : LREAL;
	LRPOSITIONPERIOD : LREAL;
END_VAR
END_FUNCTION

(* ---- L_TS2P_CALCSYNCTIME.pou ---- *)
FUNCTION L_TS2P_CALCSYNCTIME : BOOL
VAR_INPUT
	LRACTMATERIALVEL : LREAL;
	LRACCMAX : LREAL;
	LRJERKSTART : LREAL;
	LRJERKEND : LREAL;
END_VAR
VAR_OUTPUT
	LRACCTIME : LREAL;
	LRACCDIST : LREAL;
END_VAR
END_FUNCTION

(* ---- L_TS2P_CHECK_CAMREFCHANGED.pou ---- *)
FUNCTION L_TS2P_CHECK_CAMREFCHANGED : BOOL
VAR_INPUT
	CAMREFNEW : MC_CAM_REF;
	CAMREFOLD : MC_CAM_REF;
END_VAR
END_FUNCTION

(* ---- L_TS2P_CHECK_CAMREFVALID.pou ---- *)
FUNCTION L_TS2P_CHECK_CAMREFVALID : BOOL
VAR_INPUT
	CAMREF : MC_CAM_REF;
END_VAR
END_FUNCTION

(* ---- _L_MB1P_AXISCONTROLBYPOS.pou ---- *)
FUNCTION_BLOCK _L_MB1P_AXISCONTROLBYPOS
VAR_INPUT
	XENABLE : BOOL;
	LRSETPOSITION : LREAL;
	LRSETVELOCITY : LREAL;
	LRSETACCELERATION : LREAL;
	ESETVALUEMODE : L_MC1P_SetValueMode := L_MC1P_SetValueMode.Pos;
END_VAR
VAR_OUTPUT
	XBUSY : BOOL;
	XCOMMANDABORTED : BOOL;
	XERROR : BOOL;
	EERRORID : L_IE1P_Error;
	LRSETPOSOUT : LREAL;
END_VAR
VAR_IN_OUT
	AXIS : AXIS_REF;
END_VAR
VAR
	LRSETPOSITION_INT : LREAL;
	XENABLE_OLD : BOOL;
	XBUSY_OLD : BOOL;
	ESTATE : L_MB1P_States;
	MC_HALT1 : MC_HALT;
	FB_FOLLOWSETVALUES : L_MC1P_FollowSetValues;
END_VAR
END_FUNCTION_BLOCK

METHOD CALL_ERRORHANDLER
END_METHOD

METHOD CALL_FBMETHODS
END_METHOD

METHOD CALL_FB_FOLLOWSETVALUES
END_METHOD

METHOD CALL_MC_HALT
END_METHOD

METHOD CALL_MC_HALT_INPUT
END_METHOD

METHOD CALL_OUTPUT
END_METHOD

METHOD CALL_RESETCOMMANDS
END_METHOD

METHOD CALL_RESETOUTPUT
END_METHOD

METHOD CALL_STATEMACHINE
END_METHOD

METHOD CALL_S000_CYCLIC
END_METHOD

METHOD CALL_S001_INIT
END_METHOD

METHOD CALL_S002_READY
END_METHOD

METHOD CALL_S999_ERROR
END_METHOD

(* ---- _L_MB1P_AXISCONTROLBYVEL.pou ---- *)
FUNCTION_BLOCK _L_MB1P_AXISCONTROLBYVEL
VAR_INPUT
	XENABLE : BOOL;
	LRSETVELOCITY : LREAL;
END_VAR
VAR_OUTPUT
	XBUSY : BOOL;
	XCOMMANDABORTED : BOOL;
	XERROR : BOOL;
	EERRORID : L_IE1P_Error;
	LRSETVELOUT : LREAL;
END_VAR
VAR_IN_OUT
	AXIS : AXIS_REF;
END_VAR
VAR
	LRSETVELOCITY_INT : LREAL;
	XENABLE_OLD : BOOL;
	XBUSY_OLD : BOOL;
	ESTATE : L_MB1P_States;
	MC_HALT1 : MC_HALT;
	FB_FOLLOWSETVALUES : L_MC1P_FollowSetValues;
END_VAR
END_FUNCTION_BLOCK

METHOD CALL_ERRORHANDLER
END_METHOD

METHOD CALL_FBMETHODS
END_METHOD

METHOD CALL_FB_FOLLOWSETVALUES
END_METHOD

METHOD CALL_MC_HALT
END_METHOD

METHOD CALL_MC_HALT_INPUT
END_METHOD

METHOD CALL_OUTPUT
END_METHOD

METHOD CALL_RESETCOMMANDS
END_METHOD

METHOD CALL_RESETOUTPUT
END_METHOD

METHOD CALL_STATEMACHINE
END_METHOD

METHOD CALL_S000_CYCLIC
END_METHOD

METHOD CALL_S001_INIT
END_METHOD

METHOD CALL_S002_READY
END_METHOD

METHOD CALL_S999_ERROR
END_METHOD

(* ---- GLOBALTEXTLIST.pou ---- *)
FUNCTION_BLOCK GLOBALTEXTLIST
VAR
	M_TEXTLISTFILE : STRING(255);
	_STNAMESPACE : STRING;
END_VAR
END_FUNCTION_BLOCK

(* ---- L_MB1P_CHECKMODULOOVERRUN.pou ---- *)
FUNCTION_BLOCK L_MB1P_CHECKMODULOOVERRUN
VAR_INPUT
	LRSETPOS : LREAL;
	LRSETVEL : LREAL;
	LRPERIOD : LREAL;
END_VAR
VAR_OUTPUT
	XOVERRUNPOS : BOOL;
	XOVERRUNNEG : BOOL;
END_VAR
VAR
	ALRMEM : ARRAY [1..7] OF LREAL;
END_VAR
END_FUNCTION_BLOCK

METHOD CALL_CHECKMODULOOVERRUN
VAR_IN_OUT
	LRSETPOS : LREAL;
	LRSETVEL : LREAL;
	LRPERIOD : LREAL;
	XOVERRUNPOS : BOOL;
	XOVERRUNNEG : BOOL;
	ALRMEM : ARRAY [1..7] OF LREAL;
END_VAR
END_METHOD

(* ---- L_MB1P_CHECKUNLIMITEDOVERRUN.pou ---- *)
FUNCTION_BLOCK L_MB1P_CHECKUNLIMITEDOVERRUN
VAR_INPUT
	LRSETPOS : LREAL;
	LRSETVEL : LREAL;
	LRPERIOD : LREAL;
END_VAR
VAR_OUTPUT
	XOVERRUNPOS : BOOL;
	XOVERRUNNEG : BOOL;
END_VAR
VAR
	ALRMEM : ARRAY [1..7] OF LREAL;
END_VAR
END_FUNCTION_BLOCK

METHOD CALL_CHECKUNLIMITEDOVERRUN
VAR_IN_OUT
	LRSETPOS : LREAL;
	LRSETVEL : LREAL;
	LRPERIOD : LREAL;
	XOVERRUNPOS : BOOL;
	XOVERRUNNEG : BOOL;
	ALRMEM : ARRAY [1..7] OF LREAL;
END_VAR
END_METHOD

(* ---- L_MB1P_CLUTCHEXTENDEDBASE.pou ---- *)
FUNCTION_BLOCK L_MB1P_CLUTCHEXTENDEDBASE EXTENDS L_MC2P_ClutchBasic
VAR_INPUT
	XENABLE : BOOL;
	XCLUTCHCLOSE : BOOL;
	XCLUTCHOPENINSTANT : BOOL;
	ECLUTCHMODE : L_MB1P_ClutchMode := L_MB1P_ClutchMode.ramp_pos;
	ECLUTCHDIRECTION : L_MC2P_ClutchDirection := L_MC2P_ClutchDirection.mcCurrentDirection;
	EDIRECTION : L_MC1P_Direction := 0;
	LRCYCMASTERPOS : LREAL;
	LRCYCMASTERVEL : LREAL;
	LRCYCMASTERACC : LREAL;
	LRCYCSLAVEPOS : LREAL;
	LRCYCSLAVEVEL : LREAL;
	LRCYCSLAVEACC : LREAL;
	LROPENINSTANTDEC : LREAL;
	LRMASTERCLOSEPOS : LREAL;
	LRMASTERCLOSEDIST : LREAL := 100;
	LRSLAVECLOSEDIST : LREAL := 100;
	LRMASTEROPENDIST : LREAL := 100;
	LRSLAVEOPENDIST : LREAL := 100;
	LRSLAVEOPENPOS : LREAL;
	LRCLOSETIME : LREAL := 5;
	LROPENTIME : LREAL := 5;
	LRCLUTCHVEL : LREAL := 100;
	LRCLUTCHACC : LREAL := 1000.0;
	LRCLUTCHDEC : LREAL := 1000.0;
	LRCLUTCHJERK : LREAL := 1000000.0;
	LRVELTOLERANCE : LREAL := 1;
	LRAXESCYCLELENGTH : LREAL := 360;
	EMASTERTRAVERSINGRANGE : L_MC1P_TraversingRange;
	LRCYCLETIME : LREAL := 0.001;
END_VAR
VAR_OUTPUT
	XERROR : BOOL;
	EERRORID : L_IE1P_Error;
	XBUSY : BOOL;
	XDONE : BOOL;
	XSYNCHRONISED : BOOL;
	XCLUTCHACTIVE : BOOL;
	LRSETSLAVEPOSOUT : LREAL;
	LRSETSLAVEVELOUT : LREAL;
	LRSETSLAVEACCOUT : LREAL;
	LRSETSLAVEOFFSETOUT : LREAL;
	LRX0 : LREAL;
	LRX1 : LREAL;
	LRY0 : LREAL;
	LRY1 : LREAL;
	LRX0N : LREAL;
	LRX1N : LREAL;
	LRY0N : LREAL;
	LRY1N : LREAL;
	LRX0P : LREAL;
	LRX1P : LREAL;
	LRY0P : LREAL;
	LRY1P : LREAL;
END_VAR
VAR
	EAXESTRAVERSINGRANGE_INT : L_MC1P_TraversingRange;
	ECLUTCHMODE_INT : L_MB1P_ClutchMode;
	ECLUTCHDIRECTION_INT : L_MB1P_ClutchDirection;
	LRSETSLAVEOFFSET_CLUTCHREL : LREAL;
	LRSETSLAVEOFFSET_INT : LREAL;
	LRSETMASTEROFFSET_OVERRUN : LREAL;
	LRCYCLETIME_INT : LREAL;
	XCLUTCHOPENINSTANT_ACTIVE : BOOL;
	LROPENINSTANTDEC_INT : LREAL;
	XCLUTCHBASICENABLE : BOOL;
	LRTEMP : LREAL;
	LRDELTASETENDPOS : LREAL;
	LRDELTASETENDPOS_OLD : LREAL;
	LRDELTASETENDPOS_OLD2 : LREAL;
	XCLUTCHMASTERVELPOSITIVE : BOOL;
	XMASTERREVERSING : BOOL;
	XCLUTCHBASIC_EXECUTE_OLD : BOOL;
	XCLUTCHCLOSE_OLD : BOOL;
	XCLUTCHOPENINSTANT_OLD : BOOL;
	XBUSY_OLD : BOOL;
	XENABLE_OLD : BOOL;
	LRCYCMASTERPOS_OLD : LREAL;
	LRMASTERVELADD : LREAL;
	LRMASTERVELADDSYNC : LREAL;
	LRSLAVESTARTPOS : LREAL;
	LRMASTERCLOSEPOS_INT : LREAL;
	LRMASTERCLOSEDIST_INT : LREAL;
	LRSLAVECLOSEDIST_INT : LREAL;
	LRSLAVEOPENDIST_INT : LREAL;
	LRSLAVEOPENPOS_INT : LREAL;
	XSYNCMODEIN_INT : BOOL;
	LRCLUTCHTIME : LREAL;
	XCLUTCHPOSMODE_INT : BOOL := TRUE;
	LRCLUTCHVEL_INT : LREAL := 100;
	LRCLUTCHACC_INT : LREAL := 1000.0;
	LRCLUTCHDEC_INT : LREAL := 1000.0;
	LRCLUTCHJERK_INT : LREAL := 1000000.0;
	EMASTERDIRECTION_INT : L_MC2P_ClutchDirection;
	IMASTERMOVEMENTTYPE_INT : INT;
	XREVERSEALLOWED_INT : BOOL;
	XPERIODIC_INT : BOOL;
	LRSLAVEJERK : LREAL;
	ESTATE : L_MB1P_States := L_MB1P_States.INIT;
	XSTATEENTRY : BOOL;
	XSETPARAGAIN : BOOL;
	XERROR_LOCK : BOOL;
	EERRORID_LOCK : L_IE1P_Error;
	LRTOLERANCE : LREAL;
	ICYCLECNTAFTEREXECUTE : INT;
	XRESTART_INT : BOOL;
	SCCYCMASTER : L_MC2P_AxisProfile;
	SCCYCSLAVE : L_MC2P_AxisProfile;
	SCSETSLAVEOUT : L_MC2P_AxisProfile;
	SCSETSLAVEOUT_OLD : L_MC2P_AxisProfile;
	PSCSETSLAVEOUT : POINTER TO L_MC2P_AxisProfile;
	EMASTERDIRECTION : L_MC2P_ClutchDirection;
	XCLUTCHBASIC_DONE : BOOL;
	XCLUTCHBASIC_WARNINGCANTPREVENTREVERSE : BOOL;
	XCLUTCHBASIC_ERROR : BOOL;
	ECLUTCHBASIC_ERRORIDCLUTCH : L_IE1P_Error;
	XCLUTCHBASIC_BUSY : BOOL;
	XCLUTCHBASIC_CLUTCHACTIVE : BOOL;
	XCLUTCHBASIC_PERIODIC : BOOL;
	XCLUTCHBASIC_REVERSEALLOWED : BOOL;
	ECLUTCHBASIC_MASTERAXISTYPE : L_MC1P_TraversingRange;
	XCLUTCHBASIC_EXECUTE : BOOL;
	FB_CHECKMODULOOVERRUN : L_MB1P_CheckModuloOverrun;
	XHALT_OLD : BOOL;
	XHALTBUSYINT : BOOL;
	XHALTDONEINT : BOOL;
	XSIMPLEFUNRAMPSLAVEDIST : BOOL := TRUE;
	LRSETSLAVEOFFSET_CLUTCHRELENTRY : LREAL;
	XRAMPDISTABSVIALINEAR : BOOL;
	XCLUTCHBASIC_BUSY_OLD : BOOL;
	XCLUTCHMASTERVELPOSITIVE_OLD : BOOL;
	XMASTERINSIDEXSIZE : BOOL;
	XMASTERINSIDEXSIZE_OLD : BOOL;
	XMASTERINSIDEXSIZEP : BOOL;
	XMASTERINSIDEXSIZEP_OLD : BOOL;
	XMASTERINSIDEXSIZEN : BOOL;
	XMASTERINSIDEXSIZEN_OLD : BOOL;
	XCLUTCHDIRECTIONPOSITIVE : BOOL;
	ALRKOEF : ARRAY [0..5] OF LREAL;
	LRXFACTORN : LREAL;
	LRYFACTORN : LREAL;
	LRSETSLAVEOFFSET_CLUTCHRELN : LREAL;
	LRXFACTORP : LREAL;
	LRYFACTORP : LREAL;
	LRSETSLAVEOFFSET_CLUTCHRELP : LREAL;
	LRXFACTOR : LREAL;
	LRYFACTOR : LREAL;
	LRXSCALED : LREAL;
	LRYSCALED : LREAL;
	LRYSCALED_OLD : LREAL;
	LRYSCALEDDIFF : LREAL;
	LRSETYPOS : LREAL;
	LRSETYPOS_OLD : LREAL;
	LRSETYVEL : LREAL;
	LRSETYVEL_OLD : LREAL;
	LRSETYACC : LREAL;
	XCLUTCHDIRECTIONPOSITIVE_OLD : BOOL;
	LRMASTERCYCLELENGTH : LREAL;
	LRDUMMY : LREAL;
	LRCYCMASTERVEL_OLD : LREAL;
	WRAMPVELLACCSTEPPER : WORD;
	XNOREVERSEACTIVE : BOOL;
	XHALT_BUSY : BOOL;
	XHALT_DONE : BOOL;
	XSLAVEHALT : BOOL;
	C_ALRKOEF_SYNCIN : ARRAY [0..5] OF LREAL := [0, 0, 0, 1, -0.5, 0];
	C_ALRKOEF_SYNCOUT : ARRAY [0..5] OF LREAL := [0, 1, 0, -1, 0.5, 0];
END_VAR
END_FUNCTION_BLOCK

METHOD CALL_ALLOCPOINTADR
END_METHOD

METHOD CALL_CLUTCHCLOSEMODE
END_METHOD

METHOD CALL_CLUTCHOPENMODE
END_METHOD

METHOD CALL_ERRORHANDLER
END_METHOD

METHOD CALL_FBMETHODS
END_METHOD

METHOD CALL_FB_CHECKMODULOOVERRUN
END_METHOD

METHOD CALL_FB_CLUTCHBASIC
END_METHOD

METHOD CALL_FB_CLUTCHBASIC_INPUTSMASTER
END_METHOD

METHOD CALL_FB_CLUTCHBASIC_OPENINSTANT
END_METHOD

METHOD CALL_FB_CLUTCHBASIC_RAMPABS
END_METHOD

METHOD CALL_FB_CLUTCHBASIC_RAMPABS_TARGETPOS
END_METHOD

METHOD CALL_FB_CLUTCHBASIC_RAMPPOS
END_METHOD

METHOD CALL_FB_CLUTCHBASIC_RAMPREL
END_METHOD

METHOD CALL_FB_CLUTCHBASIC_RAMPSLAVEDIST
END_METHOD

METHOD CALL_FB_CLUTCHBASIC_RAMPTIME
END_METHOD

METHOD CALL_FB_CLUTCHBASIC_RAMPVELLACC
END_METHOD

METHOD CALL_FB_CLUTCHBASIC_RELATIVE
END_METHOD

METHOD CALL_MODULOTOLINEARMASTERPOS
END_METHOD

METHOD CALL_OUTPUT
END_METHOD

METHOD CALL_RAMPRELDIESTREL_CALCCOEFX0X1Y0Y1
END_METHOD

METHOD CALL_RAMPRELDISTABS_CALCCOEFX0X1Y0Y1
END_METHOD

METHOD CALL_RAMPRELDISTABS_CORRX0X1FORMODULOMASTER
END_METHOD

METHOD CALL_RAMPSLAVEDIST_ABS
END_METHOD

METHOD CALL_RAMPSLAVEDIST_REL
END_METHOD

METHOD CALL_RAMPSLAVEDIST_SETYPOSOUT
END_METHOD

METHOD CALL_RESETCLUTCH
END_METHOD

METHOD CALL_RESETCOMMANDS
END_METHOD

METHOD CALL_RESETOUTPUT
END_METHOD

METHOD CALL_SETCLUTCHCLOSEPAR
END_METHOD

METHOD CALL_SETCLUTCHCLOSEPAR_OLD
END_METHOD

METHOD CALL_SETCLUTCHOPENPAR
END_METHOD

METHOD CALL_SETCLUTCHOPENPAR_OLD
END_METHOD

METHOD CALL_STATEMASHINE
END_METHOD

METHOD SET_CLUTCHOFFSET : BOOL
VAR_INPUT
	LRIN : LREAL := 0;
END_VAR
END_METHOD

METHOD SLAVEHALT
VAR_INPUT
	XHALT : BOOL;
	SCACTSLAVE : L_MC2P_AxisProfile;
	LRMAXVELDIFF : LREAL;
	LRMAXACC : LREAL;
	LRMAXDEC : LREAL;
	LRJERK : LREAL;
	LRCYCLETIME : LREAL;
END_VAR
VAR_OUTPUT
	SCOUTPUTSLAVE : L_MC2P_AxisProfile;
	XBUSY : BOOL;
	XDONE : BOOL;
	XERROR : BOOL;
	EERRORID : L_IE1P_Error;
END_VAR
END_METHOD

METHOD CALL_S000_CYCLIC
END_METHOD

METHOD CALL_S001_INIT
END_METHOD

METHOD CALL_S010_READY
END_METHOD

METHOD CALL_S100_CLUTCH_CLOSE
END_METHOD

METHOD CALL_S200_SYNCHRON
END_METHOD

METHOD CALL_S300_CLUTCH_OPEN
END_METHOD

METHOD CALL_S998_ERROR
END_METHOD

(* ---- L_MB1P_GEARBOXPOSITION.pou ---- *)
FUNCTION_BLOCK L_MB1P_GEARBOXPOSITION EXTENDS L_MB1P_GearboxPositionBase
VAR_IN_OUT
	AXISX : AXIS_REF;
	AXISY : AXIS_REF;
END_VAR
END_FUNCTION_BLOCK

METHOD CALL_ERRORHANDLER
END_METHOD

(* ---- L_MB1P_GEARBOXPOSITIONBASE.pou ---- *)
FUNCTION_BLOCK L_MB1P_GEARBOXPOSITIONBASE
VAR_INPUT
	XENABLE : BOOL;
	LRPOSX : LREAL;
	DWNUMERATOR : DWORD := 1;
	DWDENOMINATOR : DWORD := 1;
	XLOADPOSY : BOOL;
	LRLOADPOSY : LREAL;
	LNLOADPOSYRESIDUAL : LINT;
END_VAR
VAR_OUTPUT
	LRPOSY : LREAL;
	LRVELY : LREAL;
	LNACTPOSYRESIDUAL : LINT;
	XERROR : BOOL := FALSE;
	EERRORID : L_IE1P_Error := 0;
END_VAR
VAR
	XENABLE_OLD : BOOL := FALSE;
	XINITDONE : BOOL := FALSE;
	LNPOSX : LINT := 0;
	LNPOSY : LINT := 0;
	LNPOSXOLD : LINT := 0;
	LNPOSXDIFF : LINT := 0;
	LNPOSYDIFF : LINT := 0;
	LNPOSYOLD : LINT := 0;
	LNRES_GEARBOX : LINT := 0;
	LRLENX : LREAL;
	LRLENY : LREAL;
	LRLENXOLD : LREAL;
	LRLENYOLD : LREAL;
	LRTASKCYCLE : LREAL;
	LRPOSYOLD : LREAL;
	LRGEARFACTOR : LREAL;
	DWGEARFACTOR : DWORD;
	LIAUFLOESUNG : LINT;
END_VAR
END_FUNCTION_BLOCK

METHOD CALL_S000_CYCLIC
END_METHOD

METHOD CALL_ERRORHANDLER
END_METHOD

METHOD CALL_RESET
END_METHOD

METHOD L_HLPMODULOADD : LREAL
VAR_INPUT
	LRINPUT : LINT;
	LROFFSET : LINT;
	LRLENGHT : LINT;
END_VAR
END_METHOD

METHOD L_HLPMODULODIFF : LREAL
VAR_INPUT
	LRDIFF : LINT;
	LRLEN : LINT;
END_VAR
END_METHOD

METHOD L_HLPMULDIV : LREAL
VAR_INPUT
	LNINPUT : LINT;
	DWNUMERATOR : DWORD;
	DWDENOMINATOR : DWORD;
	PLNRES : POINTER TO LINT;
END_VAR
END_METHOD

(* ---- L_MB1P_GEARBOXPOSITIONINPUT.pou ---- *)
FUNCTION_BLOCK L_MB1P_GEARBOXPOSITIONINPUT EXTENDS L_MB1P_GearboxPositionBase
VAR_INPUT
	LRCYCLELENGTHX : LREAL;
	LRCYCLELENGTHY : LREAL;
END_VAR
END_FUNCTION_BLOCK

(* ---- L_MB1P_POSPROFILERCLUTCH.pou ---- *)
FUNCTION_BLOCK L_MB1P_POSPROFILERCLUTCH
VAR_INPUT
	XENABLE : BOOL;
	XSYNCPOS : BOOL;
	XEXECUTEGAP : BOOL;
	XAUXEXECUTEGAP : BOOL;
	LRTASKCYCLETIME : LREAL := 0.001;
	LRSLAVESYNCOUTPOS : LREAL;
	LRCYCMASTERPOS : LREAL;
	LRCYCMASTERVEL : LREAL;
	LRCYCMASTERACC : LREAL;
	LRSETSLAVEPOS : LREAL;
	LRSETSLAVEVEL : LREAL;
	LRSETSLAVEACC : LREAL;
	LRJERK : LREAL := 10000;
	LRMAXACC : LREAL := 100;
	LRMAXDEC : LREAL := 100;
	LRMAXVEL : LREAL := 10;
END_VAR
VAR_OUTPUT
	XBUSY : BOOL;
	XDONE : BOOL;
	XACCDECSYNC : BOOL;
	XPOSSYNCHRONISED : BOOL;
	XERROR : BOOL;
	EERRORID : WORD;
	LRSETSLAVEPOSOUT : LREAL;
	LRSETSLAVEVELOUT : LREAL;
	LRSETSLAVEACCOUT : LREAL;
	XPROFILERESETTIMEVALID : BOOL;
	LRPROFILERESETTIME : LREAL;
END_VAR
VAR
	FB_POSPROFILERPOS : L_MC1P_PosProfiler;
	SCPROFILEPARAMETER : L_MC1P_ProfileParameter;
	WSTEPPER : WORD;
	XEXECUTEPOSPROFILER : BOOL;
	LRSLAVESYNCOUTPOS_INT : LREAL;
	XAUXEXECUTEPROFILE : BOOL;
	XEXECUTEPROFILE : BOOL;
	LRSETPOSPROFILER : LREAL;
	LRSETACCPROFILER : LREAL;
	LRSETVELPROFILER : LREAL;
	LRCYCMASTERPOS_INT : LREAL;
	LRCYCMASTERVEL_INT : LREAL;
	LRCYCMASTERACC_INT : LREAL;
	XPOSSYNCHRONISED_INT : BOOL;
	XEXECUTEGAPOLD : BOOL;
	XAUXEXECUTEGAPOLD : BOOL;
	XENABLEOLD : BOOL;
	LRCYCMASTERPOS_OLD : LREAL;
	LRTOLERANCE : LREAL;
END_VAR
END_FUNCTION_BLOCK

METHOD CALL_ERRORHANDLER
END_METHOD

METHOD CALL_FBMETHODES
END_METHOD

METHOD CALL_FB_POSPROFILERPOS
END_METHOD

METHOD CALL_FB_POSPROFILERPOSINPUTS
END_METHOD

METHOD CALL_OUTPUTS
END_METHOD

METHOD CALL_PROFILEPARAMETER
END_METHOD

METHOD CALL_RESETCOMMANDS
END_METHOD

METHOD CALL_RESETOUTPUTS
END_METHOD

METHOD CALL_STATEMACHINE
END_METHOD

(* ---- L_MB1P_POSPROFILERCLUTCHHIGH.pou ---- *)
FUNCTION_BLOCK L_MB1P_POSPROFILERCLUTCHHIGH EXTENDS L_MB1P_PosProfilerClutchState
VAR_INPUT
	XSYNCVEL : BOOL;
END_VAR
VAR_OUTPUT
	XVELSYNCHRONISED : BOOL;
END_VAR
VAR
	WSTEPPER_OLD : WORD;
	XSYNCVEL_OLD : BOOL;
	LRCYCMASTERPOSOUT : LREAL;
	LRCYCMASTERVELOUT : LREAL;
	LRCYCMASTERACCOUT : LREAL;
	LRMASTEROFFSET_INT : LREAL;
	LRSETSLAVEACCOUT_OLD : LREAL;
	LRSETSLAVEPOSOUT_OLD : LREAL;
	LRSETSLAVEPOSOUT_2OLD : LREAL;
END_VAR
END_FUNCTION_BLOCK

METHOD CALL_CALCTARGETPOS
VAR_INPUT
	LRTARGETPOS : LREAL;
END_VAR
END_METHOD

METHOD CALL_CALCLRCYCMASTERPOS
END_METHOD

METHOD CALL_OUTPUTS
END_METHOD

METHOD CALL_PROFILEPARAMETER
END_METHOD

METHOD CALL_STATEMACHINE
END_METHOD

(* ---- L_MB1P_POSPROFILERCLUTCHSTATE.pou ---- *)
FUNCTION_BLOCK L_MB1P_POSPROFILERCLUTCHSTATE EXTENDS L_MB1P_PosProfilerClutch
VAR_INPUT
	XSYNCOUTINSTANT : BOOL;
	XMOVETOTARGETPOS : BOOL;
	LRCORRECTTIMEBASE : LREAL := 0;
	LRTARGETPOS : LREAL;
	EDIRECTION : L_MC2P_ClutchDirection := L_MC2P_ClutchDirection.mcCurrentDirection;
	LRAXESCYCLELENGTH : LREAL := 360;
	EAXESTRAVERSINGRANGE : L_MC1P_TraversingRange;
	LRPOSITIONINGJERK : LREAL;
	LRPOSITIONINGACC : LREAL;
	LRPOSITIONINGDEC : LREAL;
	LRPOSITIONINGVEL : LREAL;
	LRSYNCOUTINSTANTJERK : LREAL;
	LRSYNCOUTINSTANTDEC : LREAL;
	ROVERRIDEVEL : REAL := 1.0;
	ROVERRIDEACC : REAL := 1.0;
	ROVERRIDEDEC : REAL := 1.0;
END_VAR
VAR_OUTPUT
	XREVERSING : BOOL;
	XPOSITIONING : BOOL;
	XINPOSITION : BOOL;
END_VAR
VAR
	XREVERSING_INT : BOOL;
	LRCORRECTTIMEBASE_INT : LREAL := 0;
	WMODE : WORD;
	XSYNCOUTINSTANT_OLD : BOOL;
	XMOVETOTARGETPOS_OLD : BOOL;
	XPOSMODE_INT : BOOL;
	LRTASKCYCLETIME_INT : LREAL;
	LRAXESCYCLELENGTH_INT : LREAL;
	LRTARGETPOS_INT : LREAL;
	LRTARGETPOS_LOCK : LREAL;
	LRTOLERANCEVEL : LREAL;
	LRTOLERANCEACC : LREAL;
	LRACCDIST : LREAL;
	XVELTRACE : BOOL;
	WVELTRACESTEPPER : WORD;
	LRSETACC_PROFILERPOS : LREAL;
	LRPOSPROFILERSPEED_ABS : LREAL;
	WREVERSINGVELMODE : WORD;
	LRVELZERROTOLERANZ : LREAL;
	LRSETSLAVEVELOUT_OLD : LREAL;
END_VAR
END_FUNCTION_BLOCK

METHOD CALL_CALCTARGETPOS
VAR_INPUT
	LRTARGETPOS : LREAL;
END_VAR
END_METHOD

METHOD CALL_CALCTOLERANCE
END_METHOD

METHOD CALL_CALCLRCYCMASTERPOS
END_METHOD

METHOD CALL_ERRORHANDLER
END_METHOD

METHOD CALL_FBMETHODES
END_METHOD

METHOD CALL_FB_POSPROFILERPOS
END_METHOD

METHOD CALL_FB_POSPROFILERPOSINPUTS
END_METHOD

METHOD CALL_OUTPUTS
END_METHOD

METHOD CALL_PROFILEPARAMETER
END_METHOD

METHOD CALL_PROFILEPARAMETERACCDECINMODE2
END_METHOD

METHOD CALL_RESETCOMMANDS
END_METHOD

METHOD CALL_RESETOUTPUTS
END_METHOD

METHOD CALL_STATEMACHINE
END_METHOD

(* ---- L_MB1P_STACK.pou ---- *)
FUNCTION_BLOCK L_MB1P_STACK
VAR_INPUT
	XENABLE : BOOL;
	XLOADTPPOS : BOOL;
	XLOADCYCSETPOS : BOOL;
	XTAKEPOS : BOOL;
	LRTPPOS : LREAL;
	LRCYCSETPOS : LREAL;
	LRCYCSETVEL : LREAL;
	LRPERIOD : LREAL;
	LRMINTPDIST : LREAL;
END_VAR
VAR_OUTPUT
	XBUSY : BOOL;
	XSTACKISFULL : BOOL;
	XSTACKISEMPTY : BOOL;
	LRPOSOUT : LREAL;
	LRDISTOUT : LREAL;
	LRSETDISTOUT : LREAL;
	XPOSPERIODOVERRUNPOS : BOOL;
	XPOSPERIODOVERRUNNEG : BOOL;
	UISTACKSTARTPOS : UINT := 0;
	UISTACKFILLSTATE : UINT := 0;
	ALRSTACKSAVEPOS : ARRAY [1..gc_uiStackLength] OF LREAL;
	AUIPERIODCNTRPOS : ARRAY [1..gc_uiStackLength] OF UINT;
	UIPERIODCNTR : UINT;
	LRTPDIST : LREAL;
	XPOSRECEIVED : BOOL;
	XPOSOUTOFWINDOW : BOOL;
	XWINDOWOPEN : BOOL;
END_VAR
VAR
	XSTACKVALUEVALID : BOOL;
	LRLATESTSAVEPOS : LREAL;
	UILATESTPERIODCNTRPOS : UINT;
	UICTR : UINT := 0;
	UIVARTEMP : UINT;
	XENABLE_OLD : BOOL;
	XLOADTPPOS_OLD : BOOL;
	XLOADCYCSETPOS_OLD : BOOL;
	XTAKEPOS_OLD : BOOL;
	XFIRSTLOADPOS : BOOL;
	LRCYCSETPOS_SAVE : LREAL;
	LRSETPOSDIFF : LREAL;
	XTAKEPOS_ACTIVE : BOOL;
	LRTEMPDIST : LREAL;
	LRCYCSETPOS_OLD : LREAL;
	FB_CHECKMODULOOVERRUN : L_MB1P_CheckModuloOverrun;
	GC_UISTACKLENGTH : UINT := 100;
END_VAR
END_FUNCTION_BLOCK

METHOD CALL_CNTRMODULOOVERRUN
VAR_IN_OUT
	LRCYCSETPOS : LREAL;
END_VAR
END_METHOD

METHOD CALL_FB_CHECKMODULOOVERRUN
VAR_IN_OUT
	LRCYCSETPOS : LREAL;
	LRCYCSETVEL : LREAL;
END_VAR
END_METHOD

METHOD CALL_RESETCOMMANDS
END_METHOD

METHOD CALL_RESETOUTPUT
END_METHOD

METHOD CALL_STACK
END_METHOD

METHOD CALL_STACK_LOADPOS
VAR_IN_OUT
	LRCYCPOS : LREAL;
	LRLOADPOS : LREAL;
END_VAR
END_METHOD

METHOD CALL_STACK_TAKEPOS
VAR_IN_OUT
	LRCYCPOS : LREAL;
END_VAR
END_METHOD

METHOD FUN_PERIODCNTRDIFF : LREAL
VAR_INPUT
	UIDIFF : UINT;
END_VAR
VAR_OUTPUT
	IOUT : INT;
END_VAR
END_METHOD

METHOD GET_LRLATESTDIST : LREAL
VAR_IN_OUT
	LRCYCPOS : LREAL;
END_VAR
END_METHOD

METHOD GET_LRTAKEPOS : LREAL
VAR_IN_OUT
	LRCYCPOS : LREAL;
END_VAR
END_METHOD

METHOD REVOKETAKEPOS
END_METHOD

METHOD SET_CYCSETPOS
VAR_IN_OUT
	LRCYCPOS : LREAL;
END_VAR
END_METHOD

METHOD SET_TPPOS
VAR_IN_OUT
	LRCYCPOS : LREAL;
	LRLOADTPPOS : LREAL;
END_VAR
END_METHOD

(* ---- L_MB1P_STACK_FLYINGSAW.pou ---- *)
FUNCTION_BLOCK L_MB1P_STACK_FLYINGSAW
VAR_INPUT
	XENABLE : BOOL;
	XLOADTPPOS : BOOL;
	XLOADCYCSETPOS : BOOL;
	XTAKEPOS : BOOL;
	LRTPPOS : LREAL;
	LRCYCSETPOS : LREAL;
	LRCYCSETVEL : LREAL;
	LRPERIOD : LREAL;
	LRMINTPDIST : LREAL;
END_VAR
VAR_OUTPUT
	XBUSY : BOOL;
	XSTACKISFULL : BOOL;
	XSTACKISEMPTY : BOOL;
	LRPOSOUT : LREAL;
	LRDISTOUT : LREAL;
	LRSETDISTOUT : LREAL;
	XPOSPERIODOVERRUNPOS : BOOL;
	XPOSPERIODOVERRUNNEG : BOOL;
	UISTACKSTARTPOS : UINT := 0;
	UISTACKFILLSTATE : UINT := 0;
	ALRSTACKSAVEPOS : ARRAY [1..gc_uiStackLength] OF LREAL;
	AUIPERIODCNTRPOS : ARRAY [1..gc_uiStackLength] OF UINT;
	UIPERIODCNTR : UINT;
	LRTPDIST : LREAL;
	XPOSRECEIVED : BOOL;
	XPOSOUTOFWINDOW : BOOL;
	XWINDOWOPEN : BOOL;
END_VAR
VAR
	XSTACKVALUEVALID : BOOL;
	LRLATESTSAVEPOS : LREAL;
	UILATESTPERIODCNTRPOS : UINT;
	UICTR : UINT := 0;
	UIVARTEMP : UINT;
	XENABLE_OLD : BOOL;
	XLOADTPPOS_OLD : BOOL;
	XLOADCYCSETPOS_OLD : BOOL;
	XTAKEPOS_OLD : BOOL;
	XFIRSTLOADPOS : BOOL;
	LRCYCSETPOS_SAVE : LREAL;
	LRSETPOSDIFF : LREAL;
	XTAKEPOS_ACTIVE : BOOL;
	LRTEMPDIST : LREAL;
	LRCYCSETPOS_OLD : LREAL;
	FB_CHECKMODULOOVERRUN : L_MB1P_CheckUnlimitedOverrun;
	GC_UISTACKLENGTH : UINT := 100;
END_VAR
END_FUNCTION_BLOCK

METHOD CALL_CNTRMODULOOVERRUN
VAR_IN_OUT
	LRCYCSETPOS : LREAL;
END_VAR
END_METHOD

METHOD CALL_FB_CHECKMODULOOVERRUN
VAR_IN_OUT
	LRCYCSETPOS : LREAL;
	LRCYCSETVEL : LREAL;
END_VAR
END_METHOD

METHOD CALL_RESETCOMMANDS
END_METHOD

METHOD CALL_RESETOUTPUT
END_METHOD

METHOD CALL_STACK
END_METHOD

METHOD CALL_STACK_LOADPOS
VAR_IN_OUT
	LRCYCPOS : LREAL;
	LRLOADPOS : LREAL;
END_VAR
END_METHOD

METHOD CALL_STACK_TAKEPOS
VAR_IN_OUT
	LRCYCPOS : LREAL;
END_VAR
END_METHOD

METHOD FUN_PERIODCNTRDIFF : LREAL
VAR_INPUT
	UIDIFF : UINT;
END_VAR
VAR_OUTPUT
	IOUT : INT;
END_VAR
END_METHOD

METHOD GET_LRLATESTDIST : LREAL
VAR_IN_OUT
	LRCYCPOS : LREAL;
END_VAR
END_METHOD

METHOD GET_LRTAKEPOS : LREAL
VAR_IN_OUT
	LRCYCPOS : LREAL;
END_VAR
END_METHOD

METHOD REVOKETAKEPOS
END_METHOD

METHOD SET_CYCSETPOS
VAR_IN_OUT
	LRCYCPOS : LREAL;
END_VAR
END_METHOD

METHOD SET_TPPOS
VAR_IN_OUT
	LRCYCPOS : LREAL;
	LRLOADTPPOS : LREAL;
END_VAR
END_METHOD

(* ---- L_MC2A_FINDCAMXVALUE.pou ---- *)
FUNCTION_BLOCK L_MC2A_FINDCAMXVALUE
VAR_INPUT
	LRCAMYPOSIN : LREAL;
	LRACTYPOSIN : LREAL;
	LRCYCLELENGTHX : LREAL := 360.0;
	LRCYCLELENGTHY : LREAL := 360.0;
END_VAR
VAR_OUTPUT
	LRCAMXPOSOUT : LREAL;
	LRYDIFFERENCE : LREAL;
	XBUSY : BOOL;
	XDONE : BOOL;
	XERROR : BOOL;
	EERRORID : L_IE1P_ERROR;
END_VAR
END_FUNCTION_BLOCK

METHOD METH_ADDOFFSETCYCLIC : LREAL
VAR_INPUT
	LRSETPOS : LREAL;
	LRSETOFFSET : LREAL;
	LRCYCLELENGTH : LREAL;
END_VAR
END_METHOD

METHOD METH_SHORTESTWAY : LREAL
VAR_INPUT
	LRSETPOS : LREAL;
	LRACTPOS : LREAL;
	LRCYCLELENGTH : LREAL;
END_VAR
END_METHOD

(* ---- L_TS2M_FM_FLYINGSAWSTATE.pou ---- *)
FUNCTION_BLOCK L_TS2M_FM_FLYINGSAWSTATE EXTENDS L_TB2M_FM_Base
VAR_INPUT
	ETMSTATE_EXT : L_TB2P_States;
	AXIS : REFERENCE TO AXIS_REF;
	ITFSTRUCTPROVIDER : L_TS2P_IStructProviderFlyingSaw;
	MASTERVALUES : L_MC1P_IAXIS_REF_MASTERVALUES;
	XSTARTFLYINGSAW : BOOL;
	XSYNCININSTANT : BOOL;
	XEXECUTENEXTCUT : BOOL;
	XEXECUTEGAP : BOOL;
	XSETCUTTINGLENGTHINSTANT : BOOL;
	LRCUTTINGLENGTH : LREAL;
	LRSYNCOVERRIDE : LREAL := 1;
	XSETMATERIALCOUNTER : BOOL;
	XRESUMETARGETPOS : BOOL;
	XRESETMARKSTACK : BOOL;
	PSCTPRECDATA_MARKSENSOR : POINTER TO L_MC1P.L_MC1P_TpReceiveData;
END_VAR
VAR_OUTPUT
	EFM_STATE : L_TB2P_States;
	XSYNCHRONISED : BOOL;
	XACCDECSYNC : BOOL;
	XINPOSITION : BOOL;
	XPOSITIONING : BOOL;
	LRMATERIALCOUNTER : LREAL;
	LRTARGETPOS : LREAL;
	LRCUTGAP : LREAL;
	LRACTIVECUTTINGLENGTH : LREAL;
	WMARKSINSTACK : WORD;
END_VAR
VAR
	ITFFMDATA : L_TS2M_ItfFlyingSawStateFMData := THIS^;
	ITFFLYINGSAWPROCESSING : L_TS2P_IFlyingSawProcessing := THIS^;
	MASTERVALUES_INT : L_MC1P_IAXIS_REF_MASTERVALUES;
	PDATA : POINTER TO L_TS2M_scData_FM_FlyingSaw;
	PPAR : POINTER TO L_TS2P_scPar_TM_FlyingSawState;
	PAP : POINTER TO L_TS2P_scAP_TM_FlyingSawState;
	PSF : POINTER TO L_TS2P_scSF_TM_FlyingSawState;
	FB_TRANSITION2STOPSAWERROR : L_UBUP_RequestTransitionLevel;
	FB_TRANSITION2STOPSAW : L_UBUP_RequestTransitionLevel;
	FB_TRANSITION2STARTSAW : L_UBUP_RequestTransitionEdge;
	FB_TRANSITION2STARTSAWMODECHANGE : L_UBUP_RequestTransitionEdge;
	FB_TRANSITION2SYNCINSTANT : L_UBUP_RequestTransitionEdge;
	FB_TRANSITION2SYNCLENGTHCTRLAUTO : L_UBUP_RequestTransitionLevel;
	FB_TRANSITION2SYNCLENGTHCTRLRESUME : L_UBUP_RequestTransitionEdge;
	FB_TRANSITION2SYNCMARKCTRL : L_UBUP_RequestTransitionEdge;
	FB_TRANSITION2SYNCMARKCTRLRESUME : L_UBUP_RequestTransitionEdge;
	FB_TRANSITION2SYNCSETCUTLENGTHINST : L_UBUP_RequestTransitionEdge;
	FB_TRANSITION2SYNCAFTERSYNCOUT : L_UBUP_RequestTransitionEdge;
	FB_TRANSITION2SYNCAFTERWAITING : L_UBUP_RequestTransitionLevel;
	FB_TRANSITION2SYNCFROMMOVETOLOWERLIMIT : L_UBUP_RequestTransitionEdge;
	FB_TRANSITION2SYNCFROMSYNCOUT : L_UBUP_RequestTransitionEdge;
	FB_TRANSITION2SYNCNEXTCUT : L_UBUP_RequestTransitionEdge;
	FB_TRANSITION2SYNCRESETMARKSTACK : L_UBUP_RequestTransitionEdge;
	FB_TRANSITION2SYNCOUTNEXTCUT : L_UBUP_RequestTransitionEdge;
	FB_TRANSITION2SYNCOUTRESETMARKSTACK : L_UBUP_RequestTransitionEdge;
	FB_TRANSITION2SAWSYNCHRONIZED : L_UBUP_RequestTransitionEdge;
	FB_TRANSITION2SAWSYNCHRONIZEDAFTERMOVEGAP : L_UBUP_RequestTransitionEdge;
	FB_TRANSITION2MOVETOLOWERLIMIT : L_UBUP_RequestTransitionEdge;
	FB_TRANSITION2WAITINGFORNEXTCUT : L_UBUP_RequestTransitionEdge;
	FB_TRANSITION2MOVEGAP : L_UBUP_RequestTransitionEdge;
	FB_MATERIALCOUNTER : L_TS2P_MaterialCounter;
	FB_CALCULATETARGETPOS : L_TS2P_CalculateTargetPos;
	FB_PROCESSCONTROL : L_TS2P_ProcessControl;
	FB_POSPROFILERCLUTCH : L_MB1P_PosProfilerClutchHigh;
	FB_CONTROLSETVALUES : L_MC1P_ControlSetValues;
	FB_L_TB2P_TP_CONVERTER : L_TB2P_TP_Converter;
	FB_MARKSTACK : L_TS2P_MarkStackFlyingSaw;
	FB_SYNCHRONISEDOVERRIDE : L_TS2P_SyncronisedOverride;
	FB_INPOSITION : L_TT1P_InPosition;
	FB_XEXECUTENEXTCUT_R_TRIG : R_TRIG;
	FB_XRESETMARKSTACK_R_TRIG : R_TRIG;
	XINITDONE : BOOL;
	XEXITDONE : BOOL;
	C_LRMATERIALCOUNTERCYCLELENGTH : LREAL := (16#4FFFFFFFFFFFFFFF * 1E-08);
	FLYINGSAWPROCESSING : L_TS2P_IFlyingSawProcessing;
	FMDATA : L_TS2M_ItfFlyingSawStateFMData;
	GET_LRACTIVEDEC : LREAL;
	GET_LRACTIVEJERK : LREAL;
END_VAR
END_FUNCTION_BLOCK

METHOD CALL_CALCBALANCEDPROFILE
END_METHOD

METHOD CALL_CHECKMASTERNOISE
END_METHOD

METHOD CHECKSYNCHRONISED : BOOL
END_METHOD

METHOD CALLFBS
VAR_INPUT
	ECASE : L_UBUP_StateHandleCase;
END_VAR
END_METHOD

METHOD CALLSTATE
VAR_INPUT
	ITFSTATESERVER : L_UBUP_IStateServer;
	ISTATE : INT;
	ECASE : L_UBUP_StateHandleCase;
END_VAR
END_METHOD

METHOD CHECKTRANSITION
VAR_INPUT
	ITFSTATESERVER : L_UBUP_IStateServer;
END_VAR
END_METHOD

METHOD DISABLECLIENT : BOOL
VAR_INPUT
	XFIRSTCALL : BOOL;
END_VAR
END_METHOD

METHOD ENABLECLIENT : BOOL
VAR_INPUT
	XFIRSTCALL : BOOL;
END_VAR
END_METHOD

METHOD FINALIZECYCLE
END_METHOD

METHOD LEAVESTATE
END_METHOD

METHOD PREPARECYCLE
END_METHOD

METHOD STIMULATETRANSITION
VAR_INPUT
	ECASE : L_UBUP_StateHandleCase;
END_VAR
END_METHOD

METHOD STATE_EXIT : BOOL
VAR_INPUT
	ECASE : L_UBUP_StateHandleCase;
END_VAR
END_METHOD

METHOD FB_INIT : BOOL
VAR_INPUT
	BINITRETAINS : BOOL;
	BINCOPYCODE : BOOL;
END_VAR
END_METHOD

METHOD CALL_ALLOCPOINTADR
END_METHOD

METHOD CALL_EXIT_CALLFBS
END_METHOD

METHOD CALL_MASTERAXISREF
VAR_INPUT
	MASTERVALUES : L_MC1P_IAXIS_REF_MASTERVALUES;
END_VAR
END_METHOD

METHOD CALL_RESETOUTPUT
END_METHOD

METHOD STATE_MOVE_GAP
VAR_INPUT
	ECASE : L_UBUP_StateHandleCase;
	ITFSTATESERVER : L_UBUP_IStateServer;
END_VAR
END_METHOD

METHOD STATE_MOVE_TO_LOWER_LIMIT
VAR_INPUT
	ECASE : L_UBUP_StateHandleCase;
	ITFSTATESERVER : L_UBUP_IStateServer;
END_VAR
END_METHOD

METHOD STATE_SAW_SYNCHRONIZED
VAR_INPUT
	ECASE : L_UBUP_StateHandleCase;
	ITFSTATESERVER : L_UBUP_IStateServer;
END_VAR
END_METHOD

METHOD STATE_SAW_SYNCHRONIZING
VAR_INPUT
	ECASE : L_UBUP_StateHandleCase;
	ITFSTATESERVER : L_UBUP_IStateServer;
END_VAR
END_METHOD

METHOD STATE_START_SAW
VAR_INPUT
	ECASE : L_UBUP_StateHandleCase;
	ITFSTATESERVER : L_UBUP_IStateServer;
END_VAR
END_METHOD

METHOD STATE_STOP_SAW
VAR_INPUT
	ECASE : L_UBUP_StateHandleCase;
	ITFSTATESERVER : L_UBUP_IStateServer;
END_VAR
END_METHOD

METHOD STATE_SYNC_OUT
VAR_INPUT
	ECASE : L_UBUP_StateHandleCase;
	ITFSTATESERVER : L_UBUP_IStateServer;
END_VAR
END_METHOD

METHOD STATE_WAITING_FOR_NEXT_CUT
VAR_INPUT
	ECASE : L_UBUP_StateHandleCase;
	ITFSTATESERVER : L_UBUP_IStateServer;
END_VAR
END_METHOD

METHOD CALL_FB_CALCULATETARGETPOS
END_METHOD

METHOD CALL_FB_CONTROLSETVALUES
END_METHOD

METHOD CALL_FB_INPOSITION
END_METHOD

METHOD CALL_FB_L_TB2P_TP_CONVERTER
END_METHOD

METHOD CALL_FB_MATERIALCOUNTER
END_METHOD

METHOD CALL_FB_PROCESSCONTROL
END_METHOD

METHOD CALL_FB_SYNCHRONISEDOVERRIDE
END_METHOD

METHOD TRANS_TO_SAW_SYNCHRONIZED : BOOL
END_METHOD

METHOD CLUTCH
VAR_INPUT
	ITFTECHMODULE : L_TS2P_IFlyingSawProcessing;
	XENABLE : BOOL;
	XSYNCVEL : BOOL := FALSE;
	XSYNCPOS : BOOL;
	XSYNCOUTINSTANT : BOOL;
	LRSYNCVEL : LREAL := 10;
	LRSYNCACC : LREAL := 100;
	LRSYNCDEC : LREAL := 100;
	LRSYNCJERK : LREAL := 10000;
	LRCYCMASTERPOS : LREAL;
	LRCYCMASTERVEL : LREAL;
	LRCYCMASTERACC : LREAL;
	LRSETSLAVEPOS : LREAL;
	LRSETSLAVEVEL : LREAL;
	LRSETSLAVEACC : LREAL;
END_VAR
VAR_OUTPUT
	EERRORID : L_IE1P.L_IE1P_Error;
	XERROR : BOOL;
	XBUSY : BOOL;
	XDONE : BOOL;
	XACCDECSYNC : BOOL;
	XVELSYNCHRONISED : BOOL;
	XPOSSYNCHRONISED : BOOL;
	LRSETSLAVEPOSOUT : LREAL;
	LRSETSLAVEVELOUT : LREAL;
	LRSETSLAVEACCOUT : LREAL;
	XPROFILERESETTIMEVALID : BOOL;
	LRPROFILERESETTIME : LREAL;
END_VAR
END_METHOD

METHOD EXECUTEGAP
VAR_INPUT
	ITFTECHMODULE : L_TS2P_IFlyingSawProcessing;
	XENABLE : BOOL;
	LRSYNCVEL : LREAL := 10;
	LRSYNCACC : LREAL := 100;
	LRSYNCDEC : LREAL := 100;
	LRSYNCJERK : LREAL := 10000;
	XEXECUTEGAP : BOOL;
	XAUXEXECUTEGAP : BOOL := FALSE;
	LRCYCMASTERPOS : LREAL;
	LRCYCMASTERVEL : LREAL;
	LRCYCMASTERACC : LREAL;
	LRSETSLAVEPOS : LREAL;
	LRSETSLAVEVEL : LREAL;
	LRSETSLAVEACC : LREAL;
END_VAR
VAR_OUTPUT
	EERRORID : L_IE1P.L_IE1P_Error;
	XERROR : BOOL;
	XBUSY : BOOL;
	XDONE : BOOL;
	XACCDECSYNC : BOOL;
	XVELSYNCHRONISED : BOOL;
	XPOSSYNCHRONISED : BOOL;
	LRSETSLAVEPOSOUT : LREAL;
	LRSETSLAVEVELOUT : LREAL;
	LRSETSLAVEACCOUT : LREAL;
	XPROFILERESETTIMEVALID : BOOL;
	LRPROFILERESETTIME : LREAL;
END_VAR
END_METHOD

METHOD MARKSTACK_GETMARK
VAR_INPUT
	ITFTECHMODULE : L_TS2P_IFlyingSawProcessing;
	XENABLE : BOOL;
	XGETMARK : BOOL;
	XRESETGETMARK : BOOL;
	XRESETMARKSTACK : BOOL;
	LRCYCSETPOS : LREAL;
	LRCYCSETVEL : LREAL;
END_VAR
VAR_OUTPUT
	XMARKSTACKFULL : BOOL;
	XMARKSTACKEMPTY : BOOL;
	WMARKSINSTACK : WORD;
	XMARKVALID : BOOL;
	LRMARKPOSOUT : LREAL;
END_VAR
END_METHOD

METHOD MARKSTACK_SETMARK
VAR_INPUT
	ITFTECHMODULE : L_TS2P_IFlyingSawProcessing;
	XENABLE : BOOL;
	XSETMARK : BOOL;
	LRMARKPOS : LREAL;
	XRESETMARKSTACK : BOOL;
	LRCYCSETPOS : LREAL;
	LRCYCSETVEL : LREAL;
END_VAR
VAR_OUTPUT
	XMARKSTACKFULL : BOOL;
	XMARKSTACKEMPTY : BOOL;
	WMARKSINSTACK : WORD;
	XNEWMARKRECEIVED : BOOL;
END_VAR
END_METHOD

METHOD POSITIONING
VAR_INPUT
	ITFTECHMODULE : L_TS2P_IFlyingSawProcessing;
	XENABLE : BOOL;
	XMOVETOTARGETPOS : BOOL;
	LRTARGETPOS : LREAL;
	LRPOSITIONINGVEL : LREAL;
	LRPOSITIONINGACC : LREAL;
	LRPOSITIONINGDEC : LREAL;
	LRPOSITIONINGJERK : LREAL;
	LRSETSLAVEPOS : LREAL;
	LRSETSLAVEVEL : LREAL;
	LRSETSLAVEACC : LREAL;
	LRCORRECTTIMEBASE : LREAL := 0;
	LROVERRIDE : LREAL := 1.0;
END_VAR
VAR_OUTPUT
	EERRORID : L_IE1P.L_IE1P_Error;
	XERROR : BOOL;
	XBUSY : BOOL;
	XDONE : BOOL;
	XPOSITIONING : BOOL;
	XINPOSITION : BOOL;
	LRSETSLAVEPOSOUT : LREAL;
	LRSETSLAVEVELOUT : LREAL;
	LRSETSLAVEACCOUT : LREAL;
	XPROFILERESETTIMEVALID : BOOL;
	LRPROFILERESETTIME : LREAL;
END_VAR
END_METHOD

(* ---- L_TS2M_TM_FLYINGSAWSTATE.pou ---- *)
FUNCTION_BLOCK L_TS2M_TM_FLYINGSAWSTATE EXTENDS L_TB2M_TM_MotionControl
VAR
	TM_FLYINGSAWSTATECONFIG : L_TB2P_ModuleHandlerConfig;
	PSCINPUT : POINTER TO L_TS2P_FlyingSawStateIn;
	PSCOUTPUT : POINTER TO L_TS2P_FlyingSawStateOut;
	PPAR : POINTER TO L_TS2P_scPar_TM_FlyingSawState;
	PSF : POINTER TO L_TS2P_scSF_TM_FlyingSawState;
	PAP : POINTER TO L_TS2P_scAP_TM_FlyingSawState;
	ITFTMDATA : L_TS2M_ItfFlyingSawStateTMData := THIS^;
	PDATA : POINTER TO L_TS2M_scData_FlyingSawState;
	FB_CONDDIRENABLED_SAWINPROCESS : L_UBUP_ConditionInput;
	FB_CONDDIRENABLED_MOVETOPARKPOS : L_UBUP_ConditionInput;
	FB_CONDCOLLECTSAWINPROCESS : L_UBUP_ConditionCollection := STRUCT(aitfCondition := [fb_ConditionOperationEnabled, fb_ConditionLimiter, fb_ConditionAxisHomed, fb_CondDirEnabled_SawInProcess]);
	FB_CONDCOLLECTMOVETOPARKPOS : L_UBUP_ConditionCollection := STRUCT(aitfCondition := [fb_ConditionOperationEnabled, fb_ConditionLimiter, fb_ConditionAxisHomed, fb_CondDirEnabled_MoveToParkPos]);
	FB_TRANSITION2SAWINPROCESS : L_UBUP_RequestTransitionLevel;
	FB_TRANSITION2MOVETOPARKPOS : L_UBUP_RequestTransitionEdge;
	FB_TRANSITION2MOVETOPARKPOSFROMSAWINPROCESS : L_UBUP_RequestTransitionEdge;
	FB_TRANSITION2HALTFROMSAWINPROCESS : L_UBUP_RequestTransitionEdge;
	FB_MOVETOPARKPOS : MC_MoveAbsolute;
	FB_FM_FLYINGSAW : L_TS2M_FM_FlyingSawState := STRUCT(ErrorManager := fb_ErrorManager);
	_ITFSTRUCTPROVIDERFLYINGSAW : L_TS2P_IStructProviderFlyingSaw;
	_SCTPRECEIVEDATA : L_MC1P_TpReceiveData;
	_FB_TPRECDATAPROXYMARKCORR : L_MC1P_TouchProbeRecDataProxy;
	CONNECTOR : __SYSTEM.IQueryInterface;
	FLYINGSAWPROCESSINGEXTENSION : L_TS2P_IFlyingSawProcessing;
	REMAININGTIMEOFPROFILE : LREAL;
	REMAININGTIMEOFPROFILEAVAILABLE : BOOL;
	TMDATA : L_TS2M_ItfFlyingSawStateTMData;
END_VAR
END_FUNCTION_BLOCK

METHOD CALLFBS
VAR_INPUT
	ECASE : L_UBUP_StateHandleCase;
END_VAR
END_METHOD

METHOD CALLSTATE
VAR_INPUT
	ITFSTATESERVER : L_UBUP_IStateServer;
	ISTATE : INT;
	ECASE : L_UBUP_StateHandleCase;
END_VAR
END_METHOD

METHOD CHECKTRANSITION
VAR_INPUT
	ITFSTATESERVER : L_UBUP_IStateServer;
END_VAR
END_METHOD

METHOD FINALIZECYCLE
END_METHOD

METHOD PREPARECYCLE
END_METHOD

METHOD STIMULATETRANSITION
VAR_INPUT
	ECASE : L_UBUP_StateHandleCase;
END_VAR
END_METHOD

METHOD STATE_ABORT
VAR_INPUT
	ECASE : L_UBUP_StateHandleCase;
	ITFSTATESERVER : L_UBUP_IStateServer;
END_VAR
END_METHOD

METHOD STATE_EXIT : BOOL
VAR_INPUT
	ECASE : L_UBUP_StateHandleCase;
END_VAR
END_METHOD

METHOD STATE_HALT
VAR_INPUT
	ECASE : L_UBUP_StateHandleCase;
	ITFSTATESERVER : L_UBUP_IStateServer;
END_VAR
END_METHOD

METHOD STATE_HOMING
VAR_INPUT
	ECASE : L_UBUP_StateHandleCase;
	ITFSTATESERVER : L_UBUP_IStateServer;
END_VAR
END_METHOD

METHOD STATE_MOVE_TO_PARKPOS
VAR_INPUT
	ECASE : L_UBUP_StateHandleCase;
	ITFSTATESERVER : L_UBUP_IStateServer;
END_VAR
END_METHOD

METHOD STATE_SAW_IN_PROCESS
VAR_INPUT
	ECASE : L_UBUP_StateHandleCase;
	ITFSTATESERVER : L_UBUP_IStateServer;
END_VAR
END_METHOD

METHOD STATE_STANDBY
VAR_INPUT
	ECASE : L_UBUP_StateHandleCase;
	ITFSTATESERVER : L_UBUP_IStateServer;
END_VAR
END_METHOD

METHOD CALL_ALLOCPOINTADR
END_METHOD

METHOD CALL_EXIT_CALLFBS
END_METHOD

METHOD CALL_RESETOUTPUT
END_METHOD

METHOD CALL_FM_FLYINGSAW
END_METHOD

METHOD MOVETOPARKPOS : BOOL
VAR_INPUT
	XEXECUTEMOVETOPARKPOS : BOOL;
	LRPARKPOSITION : LREAL := 180;
	EPOSITIONINGDIRECTION : MC_DIRECTION := MC_DIRECTION.mcPositiveDirection;
	LRPOSITIONINGVEL : LREAL := 10;
	LRPOSITIONINGACC : LREAL := 100;
	LRPOSITIONINGDEC : LREAL := 100;
	LRJERK : LREAL := 0;
END_VAR
VAR_OUTPUT
	XBUSY : BOOL;
	XDONE : BOOL;
	XCOMMANDABORTED : BOOL;
END_VAR
VAR_IN_OUT
	AXIS : AXIS_REF;
END_VAR
END_METHOD

(* ---- L_TS2P_ALLOWEDDIRECTION.pou ---- *)
FUNCTION_BLOCK L_TS2P_ALLOWEDDIRECTION
VAR_INPUT
	XENABLE : BOOL;
	XRESETERROR : BOOL;
	ESETVALUEMODE : L_MC1P_SetValueMode := L_MC1P_SetValueMode.Pos;
	LRSETPOSITION : LREAL;
	LRSETVELOCITY : LREAL;
	LRSETACCELERATION : LREAL;
	LRCYCLELENGTH : LREAL;
	ETRAVERSINGRANGE : L_MC1P_TraversingRange := L_MC1P_TraversingRange.Modulo;
	EALLOWEDDIRECTION : L_TB2P_AllowedDirection;
	LRALLOWEDPOSERROR : LREAL;
END_VAR
VAR_OUTPUT
	XENABLED : BOOL;
	LRSETPOSOUT : LREAL;
	LRSETVELOUT : LREAL;
	LRSETACCOUT : LREAL;
	XLIMITATIONACTIVE : BOOL;
	XWARNING : BOOL;
	XERROR : BOOL;
	EERRORID : WORD;
END_VAR
VAR
	XINITDONE : BOOL;
	LRTASKCYCLETIME : LREAL;
	LRSETPOSOUT_REVERSING : LREAL;
	XVELMODE_INT : BOOL;
	LRPOSDIFF : LREAL := 0;
	LRSETPOSDIFFINTEGRATOR : LREAL := 0;
	LRSETPOSITION_INT : LREAL;
	LRSETVELOCITY_INT : LREAL;
	LRCYCLICPOSDIFF : LREAL;
	LRSETPOSITIONOLD : LREAL;
	XMASTERINDISABLEDDIRECTION : BOOL;
	XRESETERROR_OLD : BOOL;
END_VAR
END_FUNCTION_BLOCK
